  movel([0.295404, -1.335907, -2.579843, -0.796639, 1.570796, 1.866200],accel_mss,speed_ms,0,blend_radius_m)
  movel([0.295412, -1.335943, -2.579820, -0.796627, 1.570796, 1.866208],accel_mss,speed_ms,0,blend_radius_m)
  movel([0.295403, -1.335985, -2.579792, -0.796612, 1.570796, 1.866199],accel_mss,speed_ms,0,blend_radius_m)
  movel([0.295381, -1.336040, -2.579756, -0.796593, 1.570796, 1.866177],accel_mss,speed_ms,0,blend_radius_m)
  movel([0.295349, -1.336095, -2.579721, -0.796574, 1.570796, 1.866145],accel_mss,speed_ms,0,blend_radius_m)
  movel([0.295315, -1.336133, -2.579695, -0.796560, 1.570796, 1.866112],accel_mss,speed_ms,0,blend_radius_m)
  movel([0.295270, -1.336164, -2.579675, -0.796550, 1.570796, 1.866066],accel_mss,speed_ms,0,blend_radius_m)
  movel([0.295209, -1.336190, -2.579659, -0.796541, 1.570796, 1.866006],accel_mss,speed_ms,0,blend_radius_m)
  movel([0.295150, -1.336204, -2.579649, -0.796536, 1.570796, 1.865946],accel_mss,speed_ms,0,blend_radius_m)
  movel([0.294948, -1.336225, -2.579636, -0.796528, 1.570796, 1.865745],accel_mss,speed_ms,0,blend_radius_m)
  movel([0.294564, -1.336243, -2.579624, -0.796522, 1.570796, 1.865360],accel_mss,speed_ms,0,blend_radius_m)
  movel([0.284647, -1.360640, -2.563328, -0.788421, 1.570796, 1.855443],accel_mss,speed_ms,0,blend_radius_m)
  movel([0.280975, -1.369759, -2.557027, -0.785603, 1.570796, 1.851772],accel_mss,speed_ms,0,blend_radius_m)
  movel([0.277925, -1.377354, -2.551691, -0.783344, 1.570796, 1.848721],accel_mss,speed_ms,0,blend_radius_m)
  movel([0.275199, -1.384152, -2.546846, -0.781391, 1.570796, 1.845995],accel_mss,speed_ms,0,blend_radius_m)
  movel([0.275175, -1.384193, -2.546817, -0.781379, 1.570796, 1.845972],accel_mss,speed_ms,0,blend_radius_m)
  movel([0.275139, -1.384229, -2.546791, -0.781369, 1.570796, 1.845936],accel_mss,speed_ms,0,blend_radius_m)
  speed_ms = 0.003
  movel([0.275139, -1.387342, -2.548289, -0.776758, 1.570796, 1.845936],accel_mss,speed_ms,0,blend_radius_m)
  speed_ms = 0.007
  movel([0.275100, -1.387366, -2.548271, -0.776752, 1.570796, 1.845897],accel_mss,speed_ms,0,blend_radius_m)
  movel([0.275061, -1.387375, -2.548265, -0.776749, 1.570796, 1.845858],accel_mss,speed_ms,0,blend_radius_m)
  movel([0.274454, -1.387416, -2.548235, -0.776738, 1.570796, 1.845251],accel_mss,speed_ms,0,blend_radius_m)
  movel([0.273756, -1.387452, -2.548209, -0.776728, 1.570796, 1.844552],accel_mss,speed_ms,0,blend_radius_m)
  movel([0.272946, -1.387481, -2.548189, -0.776720, 1.570796, 1.843742],accel_mss,speed_ms,0,blend_radius_m)
  movel([0.270848, -1.387542, -2.548145, -0.776703, 1.570796, 1.841644],accel_mss,speed_ms,0,blend_radius_m)
  movel([0.270977, -1.387207, -2.548386, -0.776796, 1.570796, 1.841773],accel_mss,speed_ms,0,blend_radius_m)
  movel([0.271720, -1.385272, -2.549778, -0.777339, 1.570796, 1.842517],accel_mss,speed_ms,0,blend_radius_m)
  movel([0.278710, -1.367304, -2.562451, -0.782634, 1.570796, 1.849506],accel_mss,speed_ms,0,blend_radius_m)
  movel([0.285537, -1.349959, -2.574258, -0.788172, 1.570796, 1.856333],accel_mss,speed_ms,0,blend_radius_m)
  movel([0.287626, -1.344699, -2.577757, -0.789933, 1.570796, 1.858423],accel_mss,speed_ms,0,blend_radius_m)
  movel([0.289808, -1.339211, -2.581367, -0.791811, 1.570796, 1.860604],accel_mss,speed_ms,0,blend_radius_m)
  movel([0.289826, -1.339190, -2.581381, -0.791818, 1.570796, 1.860622],accel_mss,speed_ms,0,blend_radius_m)
  movel([0.289853, -1.339171, -2.581393, -0.791825, 1.570796, 1.860650],accel_mss,speed_ms,0,blend_radius_m)
  movel([0.289881, -1.339158, -2.581402, -0.791829, 1.570796, 1.860678],accel_mss,speed_ms,0,blend_radius_m)
  movel([0.289919, -1.339144, -2.581411, -0.791834, 1.570796, 1.860715],accel_mss,speed_ms,0,blend_radius_m)
  movel([0.289955, -1.339137, -2.581415, -0.791836, 1.570796, 1.860751],accel_mss,speed_ms,0,blend_radius_m)
  movel([0.290037, -1.339134, -2.581418, -0.791838, 1.570796, 1.860833],accel_mss,speed_ms,0,blend_radius_m)
  movel([0.294408, -1.339026, -2.581488, -0.791875, 1.570796, 1.865205],accel_mss,speed_ms,0,blend_radius_m)
  movel([0.294728, -1.339025, -2.581489, -0.791875, 1.570796, 1.865524],accel_mss,speed_ms,0,blend_radius_m)
  movel([0.295043, -1.339038, -2.581480, -0.791871, 1.570796, 1.865839],accel_mss,speed_ms,0,blend_radius_m)
  movel([0.295202, -1.339055, -2.581469, -0.791865, 1.570796, 1.865998],accel_mss,speed_ms,0,blend_radius_m)
  movel([0.295351, -1.339089, -2.581447, -0.791853, 1.570796, 1.866147],accel_mss,speed_ms,0,blend_radius_m)
  movel([0.295384, -1.339105, -2.581436, -0.791847, 1.570796, 1.866180],accel_mss,speed_ms,0,blend_radius_m)
  movel([0.295404, -1.339133, -2.581418, -0.791838, 1.570796, 1.866200],accel_mss,speed_ms,0,blend_radius_m)
  movel([0.295412, -1.339168, -2.581395, -0.791826, 1.570796, 1.866208],accel_mss,speed_ms,0,blend_radius_m)
  movel([0.295403, -1.339210, -2.581368, -0.791811, 1.570796, 1.866199],accel_mss,speed_ms,0,blend_radius_m)
  movel([0.295381, -1.339266, -2.581331, -0.791792, 1.570796, 1.866177],accel_mss,speed_ms,0,blend_radius_m)
  movel([0.295349, -1.339320, -2.581296, -0.791773, 1.570796, 1.866145],accel_mss,speed_ms,0,blend_radius_m)
  movel([0.295315, -1.339358, -2.581271, -0.791760, 1.570796, 1.866112],accel_mss,speed_ms,0,blend_radius_m)
  movel([0.295270, -1.339389, -2.581251, -0.791749, 1.570796, 1.866066],accel_mss,speed_ms,0,blend_radius_m)
  movel([0.295209, -1.339415, -2.581234, -0.791740, 1.570796, 1.866006],accel_mss,speed_ms,0,blend_radius_m)
  movel([0.295150, -1.339429, -2.581224, -0.791735, 1.570796, 1.865946],accel_mss,speed_ms,0,blend_radius_m)
  movel([0.294948, -1.339450, -2.581211, -0.791728, 1.570796, 1.865745],accel_mss,speed_ms,0,blend_radius_m)
  movel([0.294564, -1.339468, -2.581199, -0.791722, 1.570796, 1.865360],accel_mss,speed_ms,0,blend_radius_m)
  movel([0.284647, -1.363810, -2.564863, -0.783716, 1.570796, 1.855443],accel_mss,speed_ms,0,blend_radius_m)
  movel([0.280975, -1.372907, -2.558548, -0.780934, 1.570796, 1.851772],accel_mss,speed_ms,0,blend_radius_m)
  movel([0.277925, -1.380483, -2.553200, -0.778706, 1.570796, 1.848721],accel_mss,speed_ms,0,blend_radius_m)
  movel([0.275199, -1.387265, -2.548344, -0.776780, 1.570796, 1.845995],accel_mss,speed_ms,0,blend_radius_m)
  movel([0.275175, -1.387306, -2.548315, -0.776768, 1.570796, 1.845972],accel_mss,speed_ms,0,blend_radius_m)
  movel([0.275139, -1.387342, -2.548289, -0.776758, 1.570796, 1.845936],accel_mss,speed_ms,0,blend_radius_m)
  speed_ms = 0.003
  movel([0.275139, -1.375017, -2.542249, -0.795123, 1.570796, 1.845936],accel_mss,speed_ms,0,blend_radius_m)
  speed_ms = 0.01
  movel([0.275139, -1.351369, -2.529790, -0.831230, 1.570796, 1.845936],accel_mss,speed_ms,0,blend_radius_m)
  movel([0.271209, -1.346627, -2.533019, -0.832743, 1.570796, 1.842006],accel_mss,speed_ms,0,blend_radius_m)
  movel([0.271209, -1.370351, -2.545537, -0.796501, 1.570796, 1.842006],accel_mss,speed_ms,0,blend_radius_m)
  speed_ms = 0.003
  movel([0.271209, -1.379596, -2.550101, -0.782692, 1.570796, 1.842006],accel_mss,speed_ms,0,blend_radius_m)
  speed_ms = 0.007
  movel([0.271117, -1.379629, -2.550077, -0.782683, 1.570796, 1.841914],accel_mss,speed_ms,0,blend_radius_m)
  movel([0.271027, -1.379649, -2.550063, -0.782677, 1.570796, 1.841823],accel_mss,speed_ms,0,blend_radius_m)
  movel([0.270594, -1.379710, -2.550019, -0.782659, 1.570796, 1.841390],accel_mss,speed_ms,0,blend_radius_m)
  movel([0.269882, -1.379801, -2.549955, -0.782633, 1.570796, 1.840679],accel_mss,speed_ms,0,blend_radius_m)
  movel([0.274743, -1.363411, -2.561425, -0.787552, 1.570796, 1.845540],accel_mss,speed_ms,0,blend_radius_m)
  movel([0.279790, -1.346600, -2.572805, -0.792984, 1.570796, 1.850586],accel_mss,speed_ms,0,blend_radius_m)
  movel([0.282065, -1.346298, -2.573006, -0.793085, 1.570796, 1.852861],accel_mss,speed_ms,0,blend_radius_m)
  movel([0.283357, -1.346133, -2.573115, -0.793141, 1.570796, 1.854153],accel_mss,speed_ms,0,blend_radius_m)
  movel([0.283649, -1.346104, -2.573135, -0.793150, 1.570796, 1.854445],accel_mss,speed_ms,0,blend_radius_m)
  movel([0.283936, -1.346085, -2.573147, -0.793157, 1.570796, 1.854732],accel_mss,speed_ms,0,blend_radius_m)
  movel([0.284087, -1.346083, -2.573149, -0.793157, 1.570796, 1.854884],accel_mss,speed_ms,0,blend_radius_m)
  movel([0.284233, -1.346093, -2.573142, -0.793154, 1.570796, 1.855029],accel_mss,speed_ms,0,blend_radius_m)
  movel([0.284260, -1.346103, -2.573135, -0.793151, 1.570796, 1.855057],accel_mss,speed_ms,0,blend_radius_m)
  movel([0.284280, -1.346123, -2.573122, -0.793144, 1.570796, 1.855077],accel_mss,speed_ms,0,blend_radius_m)
  movel([0.284288, -1.346151, -2.573103, -0.793134, 1.570796, 1.855085],accel_mss,speed_ms,0,blend_radius_m)
  movel([0.284283, -1.346184, -2.573082, -0.793124, 1.570796, 1.855079],accel_mss,speed_ms,0,blend_radius_m)
  movel([0.284233, -1.346332, -2.572983, -0.793074, 1.570796, 1.855029],accel_mss,speed_ms,0,blend_radius_m)
  movel([0.282454, -1.350866, -2.569954, -0.791569, 1.570796, 1.853250],accel_mss,speed_ms,0,blend_radius_m)
  movel([0.280494, -1.355873, -2.566576, -0.789940, 1.570796, 1.851291],accel_mss,speed_ms,0,blend_radius_m)
  movel([0.278207, -1.361736, -2.562577, -0.788076, 1.570796, 1.849003],accel_mss,speed_ms,0,blend_radius_m)
  movel([0.275917, -1.367616, -2.558519, -0.786255, 1.570796, 1.846713],accel_mss,speed_ms,0,blend_radius_m)
  movel([0.273935, -1.372723, -2.554954, -0.784711, 1.570796, 1.844731],accel_mss,speed_ms,0,blend_radius_m)
  movel([0.272258, -1.377061, -2.551899, -0.783429, 1.570796, 1.843055],accel_mss,speed_ms,0,blend_radius_m)
  movel([0.271919, -1.377934, -2.551281, -0.783175, 1.570796, 1.842716],accel_mss,speed_ms,0,blend_radius_m)
  movel([0.271351, -1.379441, -2.550211, -0.782737, 1.570796, 1.842148],accel_mss,speed_ms,0,blend_radius_m)
  movel([0.271312, -1.379512, -2.550160, -0.782717, 1.570796, 1.842108],accel_mss,speed_ms,0,blend_radius_m)
  movel([0.271281, -1.379546, -2.550136, -0.782707, 1.570796, 1.842078],accel_mss,speed_ms,0,blend_radius_m)
  movel([0.271248, -1.379574, -2.550116, -0.782699, 1.570796, 1.842044],accel_mss,speed_ms,0,blend_radius_m)
  movel([0.271209, -1.379596, -2.550101, -0.782692, 1.570796, 1.842006],accel_mss,speed_ms,0,blend_radius_m)
  speed_ms = 0.003
  movel([0.271209, -1.382720, -2.551606, -0.778063, 1.570796, 1.842006],accel_mss,speed_ms,0,blend_radius_m)
  speed_ms = 0.007
  movel([0.271117, -1.382753, -2.551582, -0.778054, 1.570796, 1.841914],accel_mss,speed_ms,0,blend_radius_m)
  movel([0.271027, -1.382773, -2.551568, -0.778048, 1.570796, 1.841823],accel_mss,speed_ms,0,blend_radius_m)
  movel([0.270594, -1.382834, -2.551524, -0.778031, 1.570796, 1.841390],accel_mss,speed_ms,0,blend_radius_m)
  movel([0.269882, -1.382924, -2.551460, -0.778005, 1.570796, 1.840679],accel_mss,speed_ms,0,blend_radius_m)
  movel([0.274743, -1.366574, -2.562956, -0.782858, 1.570796, 1.845540],accel_mss,speed_ms,0,blend_radius_m)
  movel([0.279790, -1.349802, -2.574363, -0.788224, 1.570796, 1.850586],accel_mss,speed_ms,0,blend_radius_m)
  movel([0.282065, -1.349501, -2.574564, -0.788324, 1.570796, 1.852861],accel_mss,speed_ms,0,blend_radius_m)
  movel([0.283357, -1.349336, -2.574674, -0.788379, 1.570796, 1.854153],accel_mss,speed_ms,0,blend_radius_m)
  movel([0.283649, -1.349307, -2.574694, -0.788388, 1.570796, 1.854445],accel_mss,speed_ms,0,blend_radius_m)
  movel([0.283936, -1.349288, -2.574707, -0.788395, 1.570796, 1.854732],accel_mss,speed_ms,0,blend_radius_m)
  movel([0.284087, -1.349286, -2.574708, -0.788395, 1.570796, 1.854884],accel_mss,speed_ms,0,blend_radius_m)
  movel([0.284233, -1.349296, -2.574701, -0.788392, 1.570796, 1.855029],accel_mss,speed_ms,0,blend_radius_m)
  movel([0.284260, -1.349306, -2.574694, -0.788389, 1.570796, 1.855057],accel_mss,speed_ms,0,blend_radius_m)
  movel([0.284280, -1.349326, -2.574681, -0.788382, 1.570796, 1.855077],accel_mss,speed_ms,0,blend_radius_m)
  movel([0.284288, -1.349354, -2.574662, -0.788373, 1.570796, 1.855085],accel_mss,speed_ms,0,blend_radius_m)
  movel([0.284283, -1.349386, -2.574641, -0.788362, 1.570796, 1.855079],accel_mss,speed_ms,0,blend_radius_m)
  movel([0.284233, -1.349534, -2.574542, -0.788313, 1.570796, 1.855029],accel_mss,speed_ms,0,blend_radius_m)
  movel([0.282454, -1.354058, -2.571505, -0.786826, 1.570796, 1.853250],accel_mss,speed_ms,0,blend_radius_m)
  movel([0.280494, -1.359054, -2.568119, -0.785216, 1.570796, 1.851291],accel_mss,speed_ms,0,blend_radius_m)
  movel([0.278207, -1.364903, -2.564110, -0.783376, 1.570796, 1.849003],accel_mss,speed_ms,0,blend_radius_m)
  movel([0.275917, -1.370769, -2.560043, -0.781578, 1.570796, 1.846713],accel_mss,speed_ms,0,blend_radius_m)
  movel([0.273935, -1.375864, -2.556470, -0.780055, 1.570796, 1.844731],accel_mss,speed_ms,0,blend_radius_m)
  movel([0.272258, -1.380191, -2.553408, -0.778790, 1.570796, 1.843055],accel_mss,speed_ms,0,blend_radius_m)
  movel([0.271919, -1.381062, -2.552788, -0.778539, 1.570796, 1.842716],accel_mss,speed_ms,0,blend_radius_m)
  movel([0.271351, -1.382565, -2.551716, -0.778107, 1.570796, 1.842148],accel_mss,speed_ms,0,blend_radius_m)
  movel([0.271312, -1.382637, -2.551665, -0.778087, 1.570796, 1.842108],accel_mss,speed_ms,0,blend_radius_m)
  movel([0.271281, -1.382670, -2.551641, -0.778077, 1.570796, 1.842078],accel_mss,speed_ms,0,blend_radius_m)
  movel([0.271248, -1.382698, -2.551621, -0.778069, 1.570796, 1.842044],accel_mss,speed_ms,0,blend_radius_m)
  movel([0.271209, -1.382720, -2.551606, -0.778063, 1.570796, 1.842006],accel_mss,speed_ms,0,blend_radius_m)
  speed_ms = 0.003
  movel([0.271209, -1.370351, -2.545537, -0.796501, 1.570796, 1.842006],accel_mss,speed_ms,0,blend_radius_m)
  speed_ms = 0.01
  movel([0.271209, -1.346627, -2.533019, -0.832743, 1.570796, 1.842006],accel_mss,speed_ms,0,blend_radius_m)
  movel([0.283720, -1.297614, -2.564685, -0.850089, 1.570796, 1.854516],accel_mss,speed_ms,0,blend_radius_m)
  movel([0.283720, -1.322065, -2.577821, -0.812503, 1.570796, 1.854516],accel_mss,speed_ms,0,blend_radius_m)
  speed_ms = 0.003
  movel([0.283720, -1.331626, -2.582617, -0.798146, 1.570796, 1.854516],accel_mss,speed_ms,0,blend_radius_m)
  speed_ms = 0.007
  movel([0.283274, -1.331697, -2.582572, -0.798121, 1.570796, 1.854071],accel_mss,speed_ms,0,blend_radius_m)
  movel([0.282766, -1.331776, -2.582521, -0.798093, 1.570796, 1.853563],accel_mss,speed_ms,0,blend_radius_m)
  movel([0.282165, -1.331861, -2.582466, -0.798062, 1.570796, 1.852961],accel_mss,speed_ms,0,blend_radius_m)
  movel([0.280602, -1.332079, -2.582325, -0.797985, 1.570796, 1.851398],accel_mss,speed_ms,0,blend_radius_m)
  movel([0.280741, -1.331617, -2.582623, -0.798149, 1.570796, 1.851537],accel_mss,speed_ms,0,blend_radius_m)
  movel([0.280880, -1.331154, -2.582922, -0.798313, 1.570796, 1.851676],accel_mss,speed_ms,0,blend_radius_m)
  movel([0.282316, -1.331363, -2.582787, -0.798239, 1.570796, 1.853112],accel_mss,speed_ms,0,blend_radius_m)
  movel([0.282867, -1.331445, -2.582734, -0.798210, 1.570796, 1.853663],accel_mss,speed_ms,0,blend_radius_m)
  movel([0.283328, -1.331519, -2.582686, -0.798184, 1.570796, 1.854125],accel_mss,speed_ms,0,blend_radius_m)
  movel([0.283733, -1.331590, -2.582641, -0.798158, 1.570796, 1.854530],accel_mss,speed_ms,0,blend_radius_m)
  movel([0.283741, -1.331598, -2.582635, -0.798156, 1.570796, 1.854537],accel_mss,speed_ms,0,blend_radius_m)
  movel([0.283739, -1.331610, -2.582628, -0.798151, 1.570796, 1.854536],accel_mss,speed_ms,0,blend_radius_m)
  movel([0.283720, -1.331626, -2.582617, -0.798146, 1.570796, 1.854516],accel_mss,speed_ms,0,blend_radius_m)
  speed_ms = 0.003
  movel([0.283720, -1.334861, -2.584200, -0.793328, 1.570796, 1.854516],accel_mss,speed_ms,0,blend_radius_m)
  speed_ms = 0.007
  movel([0.283274, -1.334931, -2.584154, -0.793303, 1.570796, 1.854071],accel_mss,speed_ms,0,blend_radius_m)
  movel([0.282766, -1.335010, -2.584103, -0.793275, 1.570796, 1.853563],accel_mss,speed_ms,0,blend_radius_m)
  movel([0.282165, -1.335096, -2.584048, -0.793245, 1.570796, 1.852961],accel_mss,speed_ms,0,blend_radius_m)
  movel([0.280602, -1.335313, -2.583907, -0.793169, 1.570796, 1.851398],accel_mss,speed_ms,0,blend_radius_m)
  movel([0.280741, -1.334852, -2.584206, -0.793331, 1.570796, 1.851537],accel_mss,speed_ms,0,blend_radius_m)
  movel([0.280880, -1.334390, -2.584505, -0.793494, 1.570796, 1.851676],accel_mss,speed_ms,0,blend_radius_m)
  movel([0.282316, -1.334598, -2.584370, -0.793420, 1.570796, 1.853112],accel_mss,speed_ms,0,blend_radius_m)
  movel([0.282867, -1.334681, -2.584317, -0.793391, 1.570796, 1.853663],accel_mss,speed_ms,0,blend_radius_m)
  movel([0.283328, -1.334754, -2.584269, -0.793365, 1.570796, 1.854125],accel_mss,speed_ms,0,blend_radius_m)
  movel([0.283733, -1.334825, -2.584223, -0.793341, 1.570796, 1.854530],accel_mss,speed_ms,0,blend_radius_m)
  movel([0.283741, -1.334833, -2.584218, -0.793338, 1.570796, 1.854537],accel_mss,speed_ms,0,blend_radius_m)
  movel([0.283739, -1.334845, -2.584211, -0.793334, 1.570796, 1.854536],accel_mss,speed_ms,0,blend_radius_m)
  movel([0.283720, -1.334861, -2.584200, -0.793328, 1.570796, 1.854516],accel_mss,speed_ms,0,blend_radius_m)
  speed_ms = 0.003
  movel([0.283720, -1.322065, -2.577821, -0.812503, 1.570796, 1.854516],accel_mss,speed_ms,0,blend_radius_m)
  speed_ms = 0.01
  movel([0.283720, -1.297614, -2.564685, -0.850089, 1.570796, 1.854516],accel_mss,speed_ms,0,blend_radius_m)
  movel([0.283763, -1.295871, -2.565756, -0.850763, 1.570796, 1.854559],accel_mss,speed_ms,0,blend_radius_m)
  movel([0.283763, -1.320346, -2.578913, -0.813130, 1.570796, 1.854559],accel_mss,speed_ms,0,blend_radius_m)
  speed_ms = 0.003
  movel([0.283763, -1.329917, -2.583718, -0.798754, 1.570796, 1.854559],accel_mss,speed_ms,0,blend_radius_m)
  speed_ms = 0.007
  movel([0.283665, -1.329924, -2.583714, -0.798751, 1.570796, 1.854461],accel_mss,speed_ms,0,blend_radius_m)
  movel([0.283573, -1.329918, -2.583718, -0.798754, 1.570796, 1.854369],accel_mss,speed_ms,0,blend_radius_m)
  movel([0.267806, -1.327695, -2.585144, -0.799550, 1.570796, 1.838602],accel_mss,speed_ms,0,blend_radius_m)
  movel([0.251809, -1.325748, -2.586388, -0.800254, 1.570796, 1.822605],accel_mss,speed_ms,0,blend_radius_m)
  movel([0.251761, -1.325735, -2.586396, -0.800258, 1.570796, 1.822557],accel_mss,speed_ms,0,blend_radius_m)
  movel([0.251724, -1.325709, -2.586412, -0.800268, 1.570796, 1.822521],accel_mss,speed_ms,0,blend_radius_m)
  movel([0.251715, -1.325681, -2.586430, -0.800278, 1.570796, 1.822511],accel_mss,speed_ms,0,blend_radius_m)
  movel([0.251725, -1.325645, -2.586453, -0.800291, 1.570796, 1.822521],accel_mss,speed_ms,0,blend_radius_m)
  movel([0.254190, -1.320979, -2.589413, -0.801998, 1.570796, 1.824987],accel_mss,speed_ms,0,blend_radius_m)
  movel([0.256668, -1.316306, -2.592348, -0.803735, 1.570796, 1.827464],accel_mss,speed_ms,0,blend_radius_m)
  movel([0.256713, -1.316240, -2.592389, -0.803760, 1.570796, 1.827509],accel_mss,speed_ms,0,blend_radius_m)
  movel([0.256772, -1.316177, -2.592429, -0.803784, 1.570796, 1.827569],accel_mss,speed_ms,0,blend_radius_m)
  movel([0.256793, -1.316164, -2.592437, -0.803789, 1.570796, 1.827589],accel_mss,speed_ms,0,blend_radius_m)
  movel([0.256813, -1.316160, -2.592439, -0.803790, 1.570796, 1.827610],accel_mss,speed_ms,0,blend_radius_m)
  movel([0.257759, -1.316208, -2.592409, -0.803772, 1.570796, 1.828555],accel_mss,speed_ms,0,blend_radius_m)
  movel([0.258816, -1.316268, -2.592371, -0.803750, 1.570796, 1.829612],accel_mss,speed_ms,0,blend_radius_m)
  movel([0.260062, -1.316349, -2.592321, -0.803719, 1.570796, 1.830859],accel_mss,speed_ms,0,blend_radius_m)
  movel([0.263935, -1.316628, -2.592146, -0.803615, 1.570796, 1.834731],accel_mss,speed_ms,0,blend_radius_m)
  movel([0.267792, -1.316934, -2.591955, -0.803500, 1.570796, 1.838588],accel_mss,speed_ms,0,blend_radius_m)
  movel([0.269155, -1.317054, -2.591880, -0.803455, 1.570796, 1.839952],accel_mss,speed_ms,0,blend_radius_m)
  movel([0.270512, -1.317186, -2.591797, -0.803406, 1.570796, 1.841308],accel_mss,speed_ms,0,blend_radius_m)
  movel([0.271861, -1.317333, -2.591705, -0.803351, 1.570796, 1.842657],accel_mss,speed_ms,0,blend_radius_m)
  movel([0.272781, -1.317446, -2.591634, -0.803309, 1.570796, 1.843577],accel_mss,speed_ms,0,blend_radius_m)
  movel([0.273693, -1.317576, -2.591553, -0.803260, 1.570796, 1.844489],accel_mss,speed_ms,0,blend_radius_m)
  movel([0.274595, -1.317721, -2.591462, -0.803206, 1.570796, 1.845392],accel_mss,speed_ms,0,blend_radius_m)
  movel([0.275414, -1.317867, -2.591370, -0.803152, 1.570796, 1.846211],accel_mss,speed_ms,0,blend_radius_m)
  movel([0.276222, -1.318035, -2.591265, -0.803089, 1.570796, 1.847018],accel_mss,speed_ms,0,blend_radius_m)
  movel([0.277016, -1.318219, -2.591150, -0.803021, 1.570796, 1.847813],accel_mss,speed_ms,0,blend_radius_m)
  movel([0.277714, -1.318399, -2.591036, -0.802953, 1.570796, 1.848511],accel_mss,speed_ms,0,blend_radius_m)
  movel([0.278399, -1.318598, -2.590911, -0.802879, 1.570796, 1.849196],accel_mss,speed_ms,0,blend_radius_m)
  movel([0.279071, -1.318816, -2.590774, -0.802798, 1.570796, 1.849867],accel_mss,speed_ms,0,blend_radius_m)
  movel([0.279730, -1.319051, -2.590627, -0.802711, 1.570796, 1.850526],accel_mss,speed_ms,0,blend_radius_m)
  movel([0.280376, -1.319301, -2.590469, -0.802618, 1.570796, 1.851173],accel_mss,speed_ms,0,blend_radius_m)
  movel([0.281010, -1.319571, -2.590300, -0.802518, 1.570796, 1.851806],accel_mss,speed_ms,0,blend_radius_m)
  movel([0.281379, -1.319745, -2.590190, -0.802454, 1.570796, 1.852176],accel_mss,speed_ms,0,blend_radius_m)
  movel([0.281738, -1.319934, -2.590071, -0.802384, 1.570796, 1.852534],accel_mss,speed_ms,0,blend_radius_m)
  movel([0.282081, -1.320138, -2.589943, -0.802308, 1.570796, 1.852878],accel_mss,speed_ms,0,blend_radius_m)
  movel([0.282417, -1.320353, -2.589807, -0.802229, 1.570796, 1.853213],accel_mss,speed_ms,0,blend_radius_m)
  movel([0.282735, -1.320585, -2.589661, -0.802143, 1.570796, 1.853531],accel_mss,speed_ms,0,blend_radius_m)
  movel([0.283041, -1.320830, -2.589506, -0.802052, 1.570796, 1.853838],accel_mss,speed_ms,0,blend_radius_m)
  movel([0.283334, -1.321089, -2.589343, -0.801957, 1.570796, 1.854130],accel_mss,speed_ms,0,blend_radius_m)
  movel([0.283610, -1.321359, -2.589172, -0.801857, 1.570796, 1.854407],accel_mss,speed_ms,0,blend_radius_m)
  movel([0.283835, -1.321600, -2.589020, -0.801769, 1.570796, 1.854632],accel_mss,speed_ms,0,blend_radius_m)
  movel([0.284041, -1.321857, -2.588858, -0.801674, 1.570796, 1.854837],accel_mss,speed_ms,0,blend_radius_m)
  movel([0.284233, -1.322123, -2.588690, -0.801577, 1.570796, 1.855030],accel_mss,speed_ms,0,blend_radius_m)
  movel([0.284407, -1.322403, -2.588512, -0.801474, 1.570796, 1.855203],accel_mss,speed_ms,0,blend_radius_m)
  movel([0.284568, -1.322694, -2.588328, -0.801367, 1.570796, 1.855364],accel_mss,speed_ms,0,blend_radius_m)
  movel([0.284710, -1.322997, -2.588136, -0.801256, 1.570796, 1.855506],accel_mss,speed_ms,0,blend_radius_m)
  movel([0.284835, -1.323310, -2.587938, -0.801141, 1.570796, 1.855631],accel_mss,speed_ms,0,blend_radius_m)
  movel([0.284944, -1.323634, -2.587732, -0.801023, 1.570796, 1.855740],accel_mss,speed_ms,0,blend_radius_m)
  movel([0.285032, -1.323956, -2.587528, -0.800906, 1.570796, 1.855828],accel_mss,speed_ms,0,blend_radius_m)
  movel([0.285100, -1.324285, -2.587319, -0.800785, 1.570796, 1.855897],accel_mss,speed_ms,0,blend_radius_m)
  movel([0.285151, -1.324626, -2.587102, -0.800661, 1.570796, 1.855947],accel_mss,speed_ms,0,blend_radius_m)
  movel([0.285182, -1.324974, -2.586880, -0.800535, 1.570796, 1.855979],accel_mss,speed_ms,0,blend_radius_m)
  movel([0.285194, -1.325332, -2.586653, -0.800405, 1.570796, 1.855990],accel_mss,speed_ms,0,blend_radius_m)
  movel([0.285186, -1.325696, -2.586420, -0.800272, 1.570796, 1.855982],accel_mss,speed_ms,0,blend_radius_m)
  movel([0.285163, -1.326065, -2.586185, -0.800139, 1.570796, 1.855959],accel_mss,speed_ms,0,blend_radius_m)
  movel([0.285118, -1.326442, -2.585945, -0.800002, 1.570796, 1.855914],accel_mss,speed_ms,0,blend_radius_m)
  movel([0.285089, -1.326615, -2.585834, -0.799940, 1.570796, 1.855885],accel_mss,speed_ms,0,blend_radius_m)
  movel([0.285048, -1.326789, -2.585723, -0.799877, 1.570796, 1.855844],accel_mss,speed_ms,0,blend_radius_m)
  movel([0.284996, -1.326967, -2.585609, -0.799813, 1.570796, 1.855792],accel_mss,speed_ms,0,blend_radius_m)
  movel([0.284808, -1.327550, -2.585236, -0.799602, 1.570796, 1.855605],accel_mss,speed_ms,0,blend_radius_m)
  movel([0.284614, -1.328133, -2.584863, -0.799393, 1.570796, 1.855410],accel_mss,speed_ms,0,blend_radius_m)
  movel([0.284200, -1.329332, -2.584094, -0.798963, 1.570796, 1.854997],accel_mss,speed_ms,0,blend_radius_m)
  movel([0.284152, -1.329451, -2.584018, -0.798920, 1.570796, 1.854948],accel_mss,speed_ms,0,blend_radius_m)
  movel([0.284092, -1.329568, -2.583943, -0.798879, 1.570796, 1.854889],accel_mss,speed_ms,0,blend_radius_m)
  movel([0.284020, -1.329686, -2.583867, -0.798836, 1.570796, 1.854817],accel_mss,speed_ms,0,blend_radius_m)
  movel([0.283957, -1.329768, -2.583814, -0.798807, 1.570796, 1.854753],accel_mss,speed_ms,0,blend_radius_m)
  movel([0.283884, -1.329843, -2.583766, -0.798780, 1.570796, 1.854680],accel_mss,speed_ms,0,blend_radius_m)
  movel([0.283815, -1.329896, -2.583732, -0.798761, 1.570796, 1.854611],accel_mss,speed_ms,0,blend_radius_m)
  movel([0.283789, -1.329909, -2.583723, -0.798757, 1.570796, 1.854586],accel_mss,speed_ms,0,blend_radius_m)
  movel([0.283763, -1.329917, -2.583718, -0.798754, 1.570796, 1.854559],accel_mss,speed_ms,0,blend_radius_m)
  speed_ms = 0.003
  movel([0.283763, -1.333156, -2.585304, -0.793930, 1.570796, 1.854559],accel_mss,speed_ms,0,blend_radius_m)
  speed_ms = 0.007
  movel([0.283665, -1.333162, -2.585299, -0.793927, 1.570796, 1.854461],accel_mss,speed_ms,0,blend_radius_m)
  movel([0.283573, -1.333157, -2.585303, -0.793929, 1.570796, 1.854369],accel_mss,speed_ms,0,blend_radius_m)
  movel([0.267806, -1.330938, -2.586733, -0.794718, 1.570796, 1.838602],accel_mss,speed_ms,0,blend_radius_m)
  movel([0.251809, -1.328995, -2.587980, -0.795414, 1.570796, 1.822605],accel_mss,speed_ms,0,blend_radius_m)
  movel([0.251761, -1.328983, -2.587988, -0.795418, 1.570796, 1.822557],accel_mss,speed_ms,0,blend_radius_m)
  movel([0.251724, -1.328957, -2.588005, -0.795428, 1.570796, 1.822521],accel_mss,speed_ms,0,blend_radius_m)
  movel([0.251715, -1.328929, -2.588023, -0.795438, 1.570796, 1.822511],accel_mss,speed_ms,0,blend_radius_m)
  movel([0.251725, -1.328893, -2.588046, -0.795451, 1.570796, 1.822521],accel_mss,speed_ms,0,blend_radius_m)
  movel([0.254190, -1.324237, -2.591013, -0.797140, 1.570796, 1.824987],accel_mss,speed_ms,0,blend_radius_m)
  movel([0.256668, -1.319574, -2.593956, -0.798860, 1.570796, 1.827464],accel_mss,speed_ms,0,blend_radius_m)
  movel([0.256713, -1.319508, -2.593997, -0.798884, 1.570796, 1.827509],accel_mss,speed_ms,0,blend_radius_m)
  movel([0.256772, -1.319445, -2.594037, -0.798908, 1.570796, 1.827569],accel_mss,speed_ms,0,blend_radius_m)
  movel([0.256793, -1.319432, -2.594045, -0.798913, 1.570796, 1.827589],accel_mss,speed_ms,0,blend_radius_m)
  movel([0.256813, -1.319428, -2.594047, -0.798914, 1.570796, 1.827610],accel_mss,speed_ms,0,blend_radius_m)
  movel([0.257759, -1.319476, -2.594017, -0.798896, 1.570796, 1.828555],accel_mss,speed_ms,0,blend_radius_m)
  movel([0.258816, -1.319536, -2.593979, -0.798874, 1.570796, 1.829612],accel_mss,speed_ms,0,blend_radius_m)
  movel([0.260062, -1.319616, -2.593929, -0.798844, 1.570796, 1.830859],accel_mss,speed_ms,0,blend_radius_m)
  movel([0.263935, -1.319895, -2.593754, -0.798740, 1.570796, 1.834731],accel_mss,speed_ms,0,blend_radius_m)
  movel([0.267792, -1.320200, -2.593562, -0.798627, 1.570796, 1.838588],accel_mss,speed_ms,0,blend_radius_m)
  movel([0.269155, -1.320320, -2.593486, -0.798582, 1.570796, 1.839952],accel_mss,speed_ms,0,blend_radius_m)
  movel([0.270512, -1.320452, -2.593403, -0.798533, 1.570796, 1.841308],accel_mss,speed_ms,0,blend_radius_m)
  movel([0.271861, -1.320599, -2.593311, -0.798479, 1.570796, 1.842657],accel_mss,speed_ms,0,blend_radius_m)
  movel([0.272781, -1.320711, -2.593240, -0.798438, 1.570796, 1.843577],accel_mss,speed_ms,0,blend_radius_m)
  movel([0.273693, -1.320841, -2.593158, -0.798389, 1.570796, 1.844489],accel_mss,speed_ms,0,blend_radius_m)
  movel([0.274595, -1.320986, -2.593068, -0.798336, 1.570796, 1.845392],accel_mss,speed_ms,0,blend_radius_m)
  movel([0.275414, -1.321132, -2.592975, -0.798282, 1.570796, 1.846211],accel_mss,speed_ms,0,blend_radius_m)
  movel([0.276222, -1.321299, -2.592870, -0.798220, 1.570796, 1.847018],accel_mss,speed_ms,0,blend_radius_m)
  movel([0.277016, -1.321483, -2.592754, -0.798152, 1.570796, 1.847813],accel_mss,speed_ms,0,blend_radius_m)
  movel([0.277714, -1.321663, -2.592641, -0.798086, 1.570796, 1.848511],accel_mss,speed_ms,0,blend_radius_m)
  movel([0.278399, -1.321861, -2.592515, -0.798012, 1.570796, 1.849196],accel_mss,speed_ms,0,blend_radius_m)
  movel([0.279071, -1.322079, -2.592378, -0.797932, 1.570796, 1.849867],accel_mss,speed_ms,0,blend_radius_m)
  movel([0.279730, -1.322313, -2.592230, -0.797846, 1.570796, 1.850526],accel_mss,speed_ms,0,blend_radius_m)
  movel([0.280376, -1.322563, -2.592072, -0.797754, 1.570796, 1.851173],accel_mss,speed_ms,0,blend_radius_m)
  movel([0.281010, -1.322831, -2.591903, -0.797655, 1.570796, 1.851806],accel_mss,speed_ms,0,blend_radius_m)
  movel([0.281379, -1.323006, -2.591792, -0.797591, 1.570796, 1.852176],accel_mss,speed_ms,0,blend_radius_m)
  movel([0.281738, -1.323194, -2.591673, -0.797522, 1.570796, 1.852534],accel_mss,speed_ms,0,blend_radius_m)
  movel([0.282081, -1.323398, -2.591544, -0.797447, 1.570796, 1.852878],accel_mss,speed_ms,0,blend_radius_m)
  movel([0.282417, -1.323613, -2.591408, -0.797368, 1.570796, 1.853213],accel_mss,speed_ms,0,blend_radius_m)
  movel([0.282735, -1.323844, -2.591262, -0.797283, 1.570796, 1.853531],accel_mss,speed_ms,0,blend_radius_m)
  movel([0.283041, -1.324088, -2.591107, -0.797194, 1.570796, 1.853838],accel_mss,speed_ms,0,blend_radius_m)
  movel([0.283334, -1.324347, -2.590943, -0.797099, 1.570796, 1.854130],accel_mss,speed_ms,0,blend_radius_m)
  movel([0.283610, -1.324616, -2.590772, -0.797001, 1.570796, 1.854407],accel_mss,speed_ms,0,blend_radius_m)
  movel([0.283835, -1.324856, -2.590620, -0.796913, 1.570796, 1.854632],accel_mss,speed_ms,0,blend_radius_m)
  movel([0.284041, -1.325113, -2.590457, -0.796820, 1.570796, 1.854837],accel_mss,speed_ms,0,blend_radius_m)
  movel([0.284233, -1.325378, -2.590288, -0.796723, 1.570796, 1.855030],accel_mss,speed_ms,0,blend_radius_m)
  movel([0.284407, -1.325658, -2.590110, -0.796621, 1.570796, 1.855203],accel_mss,speed_ms,0,blend_radius_m)
  movel([0.284568, -1.325949, -2.589925, -0.796515, 1.570796, 1.855364],accel_mss,speed_ms,0,blend_radius_m)
  movel([0.284710, -1.326251, -2.589733, -0.796405, 1.570796, 1.855506],accel_mss,speed_ms,0,blend_radius_m)
  movel([0.284835, -1.326563, -2.589534, -0.796292, 1.570796, 1.855631],accel_mss,speed_ms,0,blend_radius_m)
  movel([0.284944, -1.326886, -2.589328, -0.796175, 1.570796, 1.855740],accel_mss,speed_ms,0,blend_radius_m)
  movel([0.285032, -1.327207, -2.589123, -0.796059, 1.570796, 1.855828],accel_mss,speed_ms,0,blend_radius_m)
  movel([0.285100, -1.327536, -2.588913, -0.795940, 1.570796, 1.855897],accel_mss,speed_ms,0,blend_radius_m)
  movel([0.285151, -1.327876, -2.588696, -0.795817, 1.570796, 1.855947],accel_mss,speed_ms,0,blend_radius_m)
  movel([0.285182, -1.328223, -2.588474, -0.795692, 1.570796, 1.855979],accel_mss,speed_ms,0,blend_radius_m)
  movel([0.285194, -1.328580, -2.588246, -0.795563, 1.570796, 1.855990],accel_mss,speed_ms,0,blend_radius_m)
  movel([0.285186, -1.328944, -2.588013, -0.795432, 1.570796, 1.855982],accel_mss,speed_ms,0,blend_radius_m)
  movel([0.285163, -1.329312, -2.587777, -0.795300, 1.570796, 1.855959],accel_mss,speed_ms,0,blend_radius_m)
  movel([0.285118, -1.329688, -2.587536, -0.795165, 1.570796, 1.855914],accel_mss,speed_ms,0,blend_radius_m)
  movel([0.285089, -1.329861, -2.587425, -0.795103, 1.570796, 1.855885],accel_mss,speed_ms,0,blend_radius_m)
  movel([0.285048, -1.330035, -2.587314, -0.795041, 1.570796, 1.855844],accel_mss,speed_ms,0,blend_radius_m)
  movel([0.284996, -1.330213, -2.587199, -0.794977, 1.570796, 1.855792],accel_mss,speed_ms,0,blend_radius_m)
  movel([0.284808, -1.330794, -2.586826, -0.794769, 1.570796, 1.855605],accel_mss,speed_ms,0,blend_radius_m)
  movel([0.284614, -1.331376, -2.586451, -0.794562, 1.570796, 1.855410],accel_mss,speed_ms,0,blend_radius_m)
  movel([0.284200, -1.332572, -2.585681, -0.794137, 1.570796, 1.854997],accel_mss,speed_ms,0,blend_radius_m)
  movel([0.284152, -1.332691, -2.585604, -0.794094, 1.570796, 1.854948],accel_mss,speed_ms,0,blend_radius_m)
  movel([0.284092, -1.332807, -2.585529, -0.794053, 1.570796, 1.854889],accel_mss,speed_ms,0,blend_radius_m)
  movel([0.284020, -1.332925, -2.585453, -0.794011, 1.570796, 1.854817],accel_mss,speed_ms,0,blend_radius_m)
  movel([0.283957, -1.333007, -2.585400, -0.793982, 1.570796, 1.854753],accel_mss,speed_ms,0,blend_radius_m)
  movel([0.283884, -1.333082, -2.585352, -0.793956, 1.570796, 1.854680],accel_mss,speed_ms,0,blend_radius_m)
  movel([0.283815, -1.333135, -2.585317, -0.793937, 1.570796, 1.854611],accel_mss,speed_ms,0,blend_radius_m)
  movel([0.283789, -1.333147, -2.585309, -0.793932, 1.570796, 1.854586],accel_mss,speed_ms,0,blend_radius_m)
  movel([0.283763, -1.333156, -2.585304, -0.793930, 1.570796, 1.854559],accel_mss,speed_ms,0,blend_radius_m)
  speed_ms = 0.003
  movel([0.283763, -1.320346, -2.578913, -0.813130, 1.570796, 1.854559],accel_mss,speed_ms,0,blend_radius_m)
  speed_ms = 0.01
  movel([0.283763, -1.295871, -2.565756, -0.850763, 1.570796, 1.854559],accel_mss,speed_ms,0,blend_radius_m)
  movel([0.282293, -1.299239, -2.563684, -0.849465, 1.570796, 1.853089],accel_mss,speed_ms,0,blend_radius_m)
  movel([0.282293, -1.323668, -2.576799, -0.811922, 1.570796, 1.853089],accel_mss,speed_ms,0,blend_radius_m)
  speed_ms = 0.003
  movel([0.282293, -1.333219, -2.581588, -0.797582, 1.570796, 1.853089],accel_mss,speed_ms,0,blend_radius_m)
  speed_ms = 0.007
  movel([0.281918, -1.334455, -2.580786, -0.797147, 1.570796, 1.852714],accel_mss,speed_ms,0,blend_radius_m)
  movel([0.281544, -1.335690, -2.579984, -0.796715, 1.570796, 1.852341],accel_mss,speed_ms,0,blend_radius_m)
  movel([0.278441, -1.336188, -2.579660, -0.796541, 1.570796, 1.849238],accel_mss,speed_ms,0,blend_radius_m)
  movel([0.276251, -1.336569, -2.579411, -0.796409, 1.570796, 1.847047],accel_mss,speed_ms,0,blend_radius_m)
  movel([0.275394, -1.336738, -2.579301, -0.796350, 1.570796, 1.846190],accel_mss,speed_ms,0,blend_radius_m)
  movel([0.274530, -1.336932, -2.579175, -0.796282, 1.570796, 1.845326],accel_mss,speed_ms,0,blend_radius_m)
  movel([0.273708, -1.337136, -2.579041, -0.796211, 1.570796, 1.844505],accel_mss,speed_ms,0,blend_radius_m)
  movel([0.272883, -1.337362, -2.578894, -0.796133, 1.570796, 1.843679],accel_mss,speed_ms,0,blend_radius_m)
  movel([0.270940, -1.337952, -2.578508, -0.795928, 1.570796, 1.841736],accel_mss,speed_ms,0,blend_radius_m)
  movel([0.269926, -1.338289, -2.578288, -0.795812, 1.570796, 1.840722],accel_mss,speed_ms,0,blend_radius_m)
  movel([0.268912, -1.338651, -2.578052, -0.795687, 1.570796, 1.839708],accel_mss,speed_ms,0,blend_radius_m)
  movel([0.267897, -1.339034, -2.577801, -0.795555, 1.570796, 1.838694],accel_mss,speed_ms,0,blend_radius_m)
  movel([0.266884, -1.339440, -2.577535, -0.795415, 1.570796, 1.837680],accel_mss,speed_ms,0,blend_radius_m)
  movel([0.265880, -1.339865, -2.577256, -0.795268, 1.570796, 1.836676],accel_mss,speed_ms,0,blend_radius_m)
  movel([0.264877, -1.340313, -2.576961, -0.795114, 1.570796, 1.835673],accel_mss,speed_ms,0,blend_radius_m)
  movel([0.263878, -1.340784, -2.576652, -0.794953, 1.570796, 1.834675],accel_mss,speed_ms,0,blend_radius_m)
  movel([0.262881, -1.341275, -2.576329, -0.794785, 1.570796, 1.833678],accel_mss,speed_ms,0,blend_radius_m)
  movel([0.261910, -1.341780, -2.575996, -0.794613, 1.570796, 1.832706],accel_mss,speed_ms,0,blend_radius_m)
  movel([0.260943, -1.342306, -2.575650, -0.794434, 1.570796, 1.831739],accel_mss,speed_ms,0,blend_radius_m)
  movel([0.259983, -1.342850, -2.575290, -0.794248, 1.570796, 1.830780],accel_mss,speed_ms,0,blend_radius_m)
  movel([0.259028, -1.343417, -2.574916, -0.794056, 1.570796, 1.829824],accel_mss,speed_ms,0,blend_radius_m)
  movel([0.258111, -1.343985, -2.574540, -0.793864, 1.570796, 1.828907],accel_mss,speed_ms,0,blend_radius_m)
  movel([0.257201, -1.344573, -2.574150, -0.793665, 1.570796, 1.827997],accel_mss,speed_ms,0,blend_radius_m)
  movel([0.256303, -1.345181, -2.573748, -0.793461, 1.570796, 1.827100],accel_mss,speed_ms,0,blend_radius_m)
  movel([0.255412, -1.345809, -2.573331, -0.793249, 1.570796, 1.826209],accel_mss,speed_ms,0,blend_radius_m)
  movel([0.254724, -1.346319, -2.572992, -0.793078, 1.570796, 1.825520],accel_mss,speed_ms,0,blend_radius_m)
  movel([0.254047, -1.346846, -2.572641, -0.792902, 1.570796, 1.824843],accel_mss,speed_ms,0,blend_radius_m)
  movel([0.252379, -1.348218, -2.571726, -0.792445, 1.570796, 1.823175],accel_mss,speed_ms,0,blend_radius_m)
  movel([0.250748, -1.349634, -2.570780, -0.791975, 1.570796, 1.821544],accel_mss,speed_ms,0,blend_radius_m)
  movel([0.250109, -1.350216, -2.570389, -0.791783, 1.570796, 1.820906],accel_mss,speed_ms,0,blend_radius_m)
  movel([0.249486, -1.350814, -2.569988, -0.791586, 1.570796, 1.820283],accel_mss,speed_ms,0,blend_radius_m)
  movel([0.248861, -1.351441, -2.569568, -0.791380, 1.570796, 1.819657],accel_mss,speed_ms,0,blend_radius_m)
  movel([0.248252, -1.352078, -2.569139, -0.791172, 1.570796, 1.819048],accel_mss,speed_ms,0,blend_radius_m)
  movel([0.247658, -1.352723, -2.568705, -0.790961, 1.570796, 1.818454],accel_mss,speed_ms,0,blend_radius_m)
  movel([0.247081, -1.353376, -2.568265, -0.790748, 1.570796, 1.817877],accel_mss,speed_ms,0,blend_radius_m)
  movel([0.246522, -1.354036, -2.567819, -0.790534, 1.570796, 1.817318],accel_mss,speed_ms,0,blend_radius_m)
  movel([0.245984, -1.354698, -2.567372, -0.790320, 1.570796, 1.816781],accel_mss,speed_ms,0,blend_radius_m)
  movel([0.245466, -1.355366, -2.566919, -0.790104, 1.570796, 1.816263],accel_mss,speed_ms,0,blend_radius_m)
  movel([0.244966, -1.356040, -2.566463, -0.789886, 1.570796, 1.815763],accel_mss,speed_ms,0,blend_radius_m)
  movel([0.244487, -1.356719, -2.566002, -0.789668, 1.570796, 1.815283],accel_mss,speed_ms,0,blend_radius_m)
  movel([0.244025, -1.357403, -2.565537, -0.789449, 1.570796, 1.814821],accel_mss,speed_ms,0,blend_radius_m)
  movel([0.243592, -1.358077, -2.565078, -0.789234, 1.570796, 1.814388],accel_mss,speed_ms,0,blend_radius_m)
  movel([0.243180, -1.358754, -2.564616, -0.789018, 1.570796, 1.813976],accel_mss,speed_ms,0,blend_radius_m)
  movel([0.242791, -1.359434, -2.564153, -0.788803, 1.570796, 1.813587],accel_mss,speed_ms,0,blend_radius_m)
  movel([0.242421, -1.360114, -2.563688, -0.788587, 1.570796, 1.813217],accel_mss,speed_ms,0,blend_radius_m)
  movel([0.242071, -1.360799, -2.563219, -0.788371, 1.570796, 1.812867],accel_mss,speed_ms,0,blend_radius_m)
  movel([0.241755, -1.361462, -2.562765, -0.788162, 1.570796, 1.812551],accel_mss,speed_ms,0,blend_radius_m)
  movel([0.241459, -1.362128, -2.562307, -0.787953, 1.570796, 1.812256],accel_mss,speed_ms,0,blend_radius_m)
  movel([0.241191, -1.362792, -2.561852, -0.787746, 1.570796, 1.811987],accel_mss,speed_ms,0,blend_radius_m)
  movel([0.240944, -1.363453, -2.561396, -0.787539, 1.570796, 1.811740],accel_mss,speed_ms,0,blend_radius_m)
  movel([0.240721, -1.364112, -2.560942, -0.787334, 1.570796, 1.811517],accel_mss,speed_ms,0,blend_radius_m)
  movel([0.240451, -1.365015, -2.560320, -0.787055, 1.570796, 1.811247],accel_mss,speed_ms,0,blend_radius_m)
  movel([0.240217, -1.365913, -2.559699, -0.786777, 1.570796, 1.811013],accel_mss,speed_ms,0,blend_radius_m)
  movel([0.239938, -1.367112, -2.558868, -0.786409, 1.570796, 1.810734],accel_mss,speed_ms,0,blend_radius_m)
  movel([0.239680, -1.368307, -2.558038, -0.786044, 1.570796, 1.810476],accel_mss,speed_ms,0,blend_radius_m)
  movel([0.239448, -1.369472, -2.557228, -0.785690, 1.570796, 1.810244],accel_mss,speed_ms,0,blend_radius_m)
  movel([0.239237, -1.370627, -2.556422, -0.785341, 1.570796, 1.810033],accel_mss,speed_ms,0,blend_radius_m)
  movel([0.239129, -1.371375, -2.555899, -0.785115, 1.570796, 1.809925],accel_mss,speed_ms,0,blend_radius_m)
  movel([0.239064, -1.372107, -2.555386, -0.784896, 1.570796, 1.809860],accel_mss,speed_ms,0,blend_radius_m)
  movel([0.239040, -1.372671, -2.554991, -0.784727, 1.570796, 1.809837],accel_mss,speed_ms,0,blend_radius_m)
  movel([0.239038, -1.373226, -2.554601, -0.784561, 1.570796, 1.809834],accel_mss,speed_ms,0,blend_radius_m)
  movel([0.239055, -1.373774, -2.554216, -0.784398, 1.570796, 1.809852],accel_mss,speed_ms,0,blend_radius_m)
  movel([0.239094, -1.374314, -2.553837, -0.784238, 1.570796, 1.809890],accel_mss,speed_ms,0,blend_radius_m)
  movel([0.239153, -1.374844, -2.553464, -0.784081, 1.570796, 1.809949],accel_mss,speed_ms,0,blend_radius_m)
  movel([0.239230, -1.375366, -2.553096, -0.783927, 1.570796, 1.810026],accel_mss,speed_ms,0,blend_radius_m)
  movel([0.239326, -1.375877, -2.552735, -0.783777, 1.570796, 1.810122],accel_mss,speed_ms,0,blend_radius_m)
  movel([0.239469, -1.376486, -2.552305, -0.783598, 1.570796, 1.810266],accel_mss,speed_ms,0,blend_radius_m)
  movel([0.239636, -1.377085, -2.551881, -0.783422, 1.570796, 1.810432],accel_mss,speed_ms,0,blend_radius_m)
  movel([0.239830, -1.377667, -2.551470, -0.783252, 1.570796, 1.810626],accel_mss,speed_ms,0,blend_radius_m)
  movel([0.240045, -1.378236, -2.551066, -0.783087, 1.570796, 1.810841],accel_mss,speed_ms,0,blend_radius_m)
  movel([0.240284, -1.378789, -2.550674, -0.782926, 1.570796, 1.811081],accel_mss,speed_ms,0,blend_radius_m)
  movel([0.240546, -1.379327, -2.550292, -0.782770, 1.570796, 1.811342],accel_mss,speed_ms,0,blend_radius_m)
  movel([0.240841, -1.379866, -2.549908, -0.782614, 1.570796, 1.811637],accel_mss,speed_ms,0,blend_radius_m)
  movel([0.241158, -1.380389, -2.549536, -0.782464, 1.570796, 1.811955],accel_mss,speed_ms,0,blend_radius_m)
  movel([0.241499, -1.380894, -2.549177, -0.782319, 1.570796, 1.812295],accel_mss,speed_ms,0,blend_radius_m)
  movel([0.241860, -1.381384, -2.548827, -0.782178, 1.570796, 1.812657],accel_mss,speed_ms,0,blend_radius_m)
  movel([0.242243, -1.381854, -2.548491, -0.782044, 1.570796, 1.813039],accel_mss,speed_ms,0,blend_radius_m)
  movel([0.242648, -1.382308, -2.548167, -0.781914, 1.570796, 1.813444],accel_mss,speed_ms,0,blend_radius_m)
  movel([0.243080, -1.382749, -2.547851, -0.781788, 1.570796, 1.813877],accel_mss,speed_ms,0,blend_radius_m)
  movel([0.243531, -1.383173, -2.547548, -0.781668, 1.570796, 1.814327],accel_mss,speed_ms,0,blend_radius_m)
  movel([0.244002, -1.383579, -2.547257, -0.781553, 1.570796, 1.814798],accel_mss,speed_ms,0,blend_radius_m)
  movel([0.244493, -1.383965, -2.546980, -0.781443, 1.570796, 1.815290],accel_mss,speed_ms,0,blend_radius_m)
  movel([0.245003, -1.384334, -2.546716, -0.781339, 1.570796, 1.815799],accel_mss,speed_ms,0,blend_radius_m)
  movel([0.245528, -1.384683, -2.546465, -0.781241, 1.570796, 1.816325],accel_mss,speed_ms,0,blend_radius_m)
  movel([0.246115, -1.385035, -2.546212, -0.781142, 1.570796, 1.816911],accel_mss,speed_ms,0,blend_radius_m)
  movel([0.246714, -1.385368, -2.545973, -0.781048, 1.570796, 1.817511],accel_mss,speed_ms,0,blend_radius_m)
  movel([0.247335, -1.385679, -2.545749, -0.780961, 1.570796, 1.818132],accel_mss,speed_ms,0,blend_radius_m)
  movel([0.247973, -1.385969, -2.545540, -0.780880, 1.570796, 1.818769],accel_mss,speed_ms,0,blend_radius_m)
  movel([0.248627, -1.386238, -2.545347, -0.780804, 1.570796, 1.819423],accel_mss,speed_ms,0,blend_radius_m)
  movel([0.249299, -1.386484, -2.545170, -0.780736, 1.570796, 1.820095],accel_mss,speed_ms,0,blend_radius_m)
  movel([0.250013, -1.386719, -2.545000, -0.780670, 1.570796, 1.820810],accel_mss,speed_ms,0,blend_radius_m)
  movel([0.250744, -1.386937, -2.544843, -0.780609, 1.570796, 1.821540],accel_mss,speed_ms,0,blend_radius_m)
  movel([0.251487, -1.387134, -2.544701, -0.780555, 1.570796, 1.822283],accel_mss,speed_ms,0,blend_radius_m)
  movel([0.252244, -1.387308, -2.544575, -0.780506, 1.570796, 1.823041],accel_mss,speed_ms,0,blend_radius_m)
  movel([0.253013, -1.387464, -2.544462, -0.780463, 1.570796, 1.823810],accel_mss,speed_ms,0,blend_radius_m)
  movel([0.253794, -1.387601, -2.544363, -0.780425, 1.570796, 1.824591],accel_mss,speed_ms,0,blend_radius_m)
  movel([0.254605, -1.387719, -2.544278, -0.780392, 1.570796, 1.825401],accel_mss,speed_ms,0,blend_radius_m)
  movel([0.255429, -1.387815, -2.544209, -0.780365, 1.570796, 1.826225],accel_mss,speed_ms,0,blend_radius_m)
  movel([0.256261, -1.387893, -2.544152, -0.780344, 1.570796, 1.827058],accel_mss,speed_ms,0,blend_radius_m)
  movel([0.257105, -1.387950, -2.544111, -0.780328, 1.570796, 1.827901],accel_mss,speed_ms,0,blend_radius_m)
  movel([0.257958, -1.387985, -2.544086, -0.780318, 1.570796, 1.828755],accel_mss,speed_ms,0,blend_radius_m)
  movel([0.258821, -1.388002, -2.544073, -0.780313, 1.570796, 1.829617],accel_mss,speed_ms,0,blend_radius_m)
  movel([0.259693, -1.387996, -2.544078, -0.780315, 1.570796, 1.830489],accel_mss,speed_ms,0,blend_radius_m)
  movel([0.260575, -1.387970, -2.544097, -0.780322, 1.570796, 1.831371],accel_mss,speed_ms,0,blend_radius_m)
  movel([0.261462, -1.387925, -2.544129, -0.780335, 1.570796, 1.832259],accel_mss,speed_ms,0,blend_radius_m)
  movel([0.262358, -1.387858, -2.544178, -0.780353, 1.570796, 1.833154],accel_mss,speed_ms,0,blend_radius_m)
  movel([0.263262, -1.387770, -2.544241, -0.780378, 1.570796, 1.834059],accel_mss,speed_ms,0,blend_radius_m)
  movel([0.264172, -1.387663, -2.544319, -0.780407, 1.570796, 1.834968],accel_mss,speed_ms,0,blend_radius_m)
  movel([0.266174, -1.387406, -2.544504, -0.780479, 1.570796, 1.836970],accel_mss,speed_ms,0,blend_radius_m)
  movel([0.265950, -1.388175, -2.543948, -0.780265, 1.570796, 1.836746],accel_mss,speed_ms,0,blend_radius_m)
  movel([0.265726, -1.388944, -2.543392, -0.780053, 1.570796, 1.836522],accel_mss,speed_ms,0,blend_radius_m)
  movel([0.244685, -1.391802, -2.541316, -0.779271, 1.570796, 1.815481],accel_mss,speed_ms,0,blend_radius_m)
  movel([0.223610, -1.395032, -2.538956, -0.778401, 1.570796, 1.794406],accel_mss,speed_ms,0,blend_radius_m)
  movel([0.230335, -1.368198, -2.558114, -0.786077, 1.570796, 1.801132],accel_mss,speed_ms,0,blend_radius_m)
  movel([0.237492, -1.340228, -2.577017, -0.795144, 1.570796, 1.808288],accel_mss,speed_ms,0,blend_radius_m)
  movel([0.259913, -1.336512, -2.579449, -0.796428, 1.570796, 1.830709],accel_mss,speed_ms,0,blend_radius_m)
  movel([0.282293, -1.333219, -2.581588, -0.797582, 1.570796, 1.853089],accel_mss,speed_ms,0,blend_radius_m)
  speed_ms = 0.003
  movel([0.282293, -1.336450, -2.583168, -0.792771, 1.570796, 1.853089],accel_mss,speed_ms,0,blend_radius_m)
  speed_ms = 0.007
  movel([0.281918, -1.337684, -2.582364, -0.792340, 1.570796, 1.852714],accel_mss,speed_ms,0,blend_radius_m)
  movel([0.281544, -1.338916, -2.581560, -0.791913, 1.570796, 1.852341],accel_mss,speed_ms,0,blend_radius_m)
  movel([0.278441, -1.339413, -2.581235, -0.791741, 1.570796, 1.849238],accel_mss,speed_ms,0,blend_radius_m)
  movel([0.276251, -1.339793, -2.580986, -0.791610, 1.570796, 1.847047],accel_mss,speed_ms,0,blend_radius_m)
  movel([0.275394, -1.339962, -2.580875, -0.791551, 1.570796, 1.846190],accel_mss,speed_ms,0,blend_radius_m)
  movel([0.274530, -1.340156, -2.580749, -0.791485, 1.570796, 1.845326],accel_mss,speed_ms,0,blend_radius_m)
  movel([0.273708, -1.340359, -2.580615, -0.791415, 1.570796, 1.844505],accel_mss,speed_ms,0,blend_radius_m)
  movel([0.272883, -1.340584, -2.580467, -0.791337, 1.570796, 1.843679],accel_mss,speed_ms,0,blend_radius_m)
  movel([0.270940, -1.341174, -2.580081, -0.791135, 1.570796, 1.841736],accel_mss,speed_ms,0,blend_radius_m)
  movel([0.269926, -1.341509, -2.579860, -0.791020, 1.570796, 1.840722],accel_mss,speed_ms,0,blend_radius_m)
  movel([0.268912, -1.341870, -2.579623, -0.790896, 1.570796, 1.839708],accel_mss,speed_ms,0,blend_radius_m)
  movel([0.267897, -1.342252, -2.579371, -0.790765, 1.570796, 1.838694],accel_mss,speed_ms,0,blend_radius_m)
  movel([0.266884, -1.342657, -2.579105, -0.790627, 1.570796, 1.837680],accel_mss,speed_ms,0,blend_radius_m)
  movel([0.265880, -1.343082, -2.578825, -0.790482, 1.570796, 1.836676],accel_mss,speed_ms,0,blend_radius_m)
  movel([0.264877, -1.343529, -2.578530, -0.790330, 1.570796, 1.835673],accel_mss,speed_ms,0,blend_radius_m)
  movel([0.263878, -1.343999, -2.578220, -0.790171, 1.570796, 1.834675],accel_mss,speed_ms,0,blend_radius_m)
  movel([0.262881, -1.344489, -2.577896, -0.790005, 1.570796, 1.833678],accel_mss,speed_ms,0,blend_radius_m)
  movel([0.261910, -1.344993, -2.577562, -0.789834, 1.570796, 1.832706],accel_mss,speed_ms,0,blend_radius_m)
  movel([0.260943, -1.345517, -2.577215, -0.789657, 1.570796, 1.831739],accel_mss,speed_ms,0,blend_radius_m)
  movel([0.259983, -1.346061, -2.576855, -0.789474, 1.570796, 1.830780],accel_mss,speed_ms,0,blend_radius_m)
  movel([0.259028, -1.346626, -2.576479, -0.789284, 1.570796, 1.829824],accel_mss,speed_ms,0,blend_radius_m)
  movel([0.258111, -1.347192, -2.576103, -0.789094, 1.570796, 1.828907],accel_mss,speed_ms,0,blend_radius_m)
  movel([0.257201, -1.347780, -2.575712, -0.788897, 1.570796, 1.827997],accel_mss,speed_ms,0,blend_radius_m)
  movel([0.256303, -1.348386, -2.575308, -0.788695, 1.570796, 1.827100],accel_mss,speed_ms,0,blend_radius_m)
  movel([0.255412, -1.349012, -2.574890, -0.788486, 1.570796, 1.826209],accel_mss,speed_ms,0,blend_radius_m)
  movel([0.254724, -1.349521, -2.574551, -0.788317, 1.570796, 1.825520],accel_mss,speed_ms,0,blend_radius_m)
  movel([0.254047, -1.350047, -2.574199, -0.788143, 1.570796, 1.824843],accel_mss,speed_ms,0,blend_radius_m)
  movel([0.252379, -1.351416, -2.573282, -0.787691, 1.570796, 1.823175],accel_mss,speed_ms,0,blend_radius_m)
  movel([0.250748, -1.352829, -2.572333, -0.787227, 1.570796, 1.821544],accel_mss,speed_ms,0,blend_radius_m)
  movel([0.250109, -1.353410, -2.571942, -0.787037, 1.570796, 1.820906],accel_mss,speed_ms,0,blend_radius_m)
  movel([0.249486, -1.354006, -2.571540, -0.786843, 1.570796, 1.820283],accel_mss,speed_ms,0,blend_radius_m)
  movel([0.248861, -1.354631, -2.571118, -0.786639, 1.570796, 1.819657],accel_mss,speed_ms,0,blend_radius_m)
  movel([0.248252, -1.355267, -2.570689, -0.786433, 1.570796, 1.819048],accel_mss,speed_ms,0,blend_radius_m)
  movel([0.247658, -1.355910, -2.570253, -0.786225, 1.570796, 1.818454],accel_mss,speed_ms,0,blend_radius_m)
  movel([0.247081, -1.356562, -2.569812, -0.786015, 1.570796, 1.817877],accel_mss,speed_ms,0,blend_radius_m)
  movel([0.246522, -1.357221, -2.569365, -0.785803, 1.570796, 1.817318],accel_mss,speed_ms,0,blend_radius_m)
  movel([0.245984, -1.357881, -2.568917, -0.785591, 1.570796, 1.816781],accel_mss,speed_ms,0,blend_radius_m)
  movel([0.245466, -1.358548, -2.568464, -0.785378, 1.570796, 1.816263],accel_mss,speed_ms,0,blend_radius_m)
  movel([0.244966, -1.359220, -2.568006, -0.785163, 1.570796, 1.815763],accel_mss,speed_ms,0,blend_radius_m)
  movel([0.244487, -1.359897, -2.567544, -0.784948, 1.570796, 1.815283],accel_mss,speed_ms,0,blend_radius_m)
  movel([0.244025, -1.360580, -2.567078, -0.784732, 1.570796, 1.814821],accel_mss,speed_ms,0,blend_radius_m)
  movel([0.243592, -1.361253, -2.566618, -0.784519, 1.570796, 1.814388],accel_mss,speed_ms,0,blend_radius_m)
  movel([0.243180, -1.361928, -2.566155, -0.784306, 1.570796, 1.813976],accel_mss,speed_ms,0,blend_radius_m)
  movel([0.242791, -1.362606, -2.565690, -0.784093, 1.570796, 1.813587],accel_mss,speed_ms,0,blend_radius_m)
  movel([0.242421, -1.363284, -2.565224, -0.783880, 1.570796, 1.813217],accel_mss,speed_ms,0,blend_radius_m)
  movel([0.242071, -1.363968, -2.564755, -0.783667, 1.570796, 1.812867],accel_mss,speed_ms,0,blend_radius_m)
  movel([0.241755, -1.364630, -2.564299, -0.783461, 1.570796, 1.812551],accel_mss,speed_ms,0,blend_radius_m)
  movel([0.241459, -1.365294, -2.563841, -0.783254, 1.570796, 1.812256],accel_mss,speed_ms,0,blend_radius_m)
  movel([0.241191, -1.365956, -2.563384, -0.783049, 1.570796, 1.811987],accel_mss,speed_ms,0,blend_radius_m)
  movel([0.240944, -1.366616, -2.562927, -0.782846, 1.570796, 1.811740],accel_mss,speed_ms,0,blend_radius_m)
  movel([0.240721, -1.367274, -2.562472, -0.782643, 1.570796, 1.811517],accel_mss,speed_ms,0,blend_radius_m)
  movel([0.240451, -1.368174, -2.561848, -0.782367, 1.570796, 1.811247],accel_mss,speed_ms,0,blend_radius_m)
  movel([0.240217, -1.369070, -2.561226, -0.782093, 1.570796, 1.811013],accel_mss,speed_ms,0,blend_radius_m)
  movel([0.239938, -1.370267, -2.560393, -0.781730, 1.570796, 1.810734],accel_mss,speed_ms,0,blend_radius_m)
  movel([0.239680, -1.371458, -2.559561, -0.781369, 1.570796, 1.810476],accel_mss,speed_ms,0,blend_radius_m)
  movel([0.239448, -1.372620, -2.558749, -0.781020, 1.570796, 1.810244],accel_mss,speed_ms,0,blend_radius_m)
  movel([0.239237, -1.373773, -2.557941, -0.780675, 1.570796, 1.810033],accel_mss,speed_ms,0,blend_radius_m)
  movel([0.239129, -1.374519, -2.557417, -0.780453, 1.570796, 1.809925],accel_mss,speed_ms,0,blend_radius_m)
  movel([0.239064, -1.375249, -2.556903, -0.780236, 1.570796, 1.809860],accel_mss,speed_ms,0,blend_radius_m)
  movel([0.239040, -1.375811, -2.556507, -0.780070, 1.570796, 1.809837],accel_mss,speed_ms,0,blend_radius_m)
  movel([0.239038, -1.376366, -2.556117, -0.779907, 1.570796, 1.809834],accel_mss,speed_ms,0,blend_radius_m)
  movel([0.239055, -1.376912, -2.555731, -0.779746, 1.570796, 1.809852],accel_mss,speed_ms,0,blend_radius_m)
  movel([0.239094, -1.377451, -2.555350, -0.779588, 1.570796, 1.809890],accel_mss,speed_ms,0,blend_radius_m)
  movel([0.239153, -1.377979, -2.554976, -0.779433, 1.570796, 1.809949],accel_mss,speed_ms,0,blend_radius_m)
  movel([0.239230, -1.378501, -2.554607, -0.779281, 1.570796, 1.810026],accel_mss,speed_ms,0,blend_radius_m)
  movel([0.239326, -1.379010, -2.554246, -0.779133, 1.570796, 1.810122],accel_mss,speed_ms,0,blend_radius_m)
  movel([0.239469, -1.379618, -2.553815, -0.778956, 1.570796, 1.810266],accel_mss,speed_ms,0,blend_radius_m)
  movel([0.239636, -1.380216, -2.553390, -0.778783, 1.570796, 1.810432],accel_mss,speed_ms,0,blend_radius_m)
  movel([0.239830, -1.380796, -2.552978, -0.778615, 1.570796, 1.810626],accel_mss,speed_ms,0,blend_radius_m)
  movel([0.240045, -1.381364, -2.552573, -0.778452, 1.570796, 1.810841],accel_mss,speed_ms,0,blend_radius_m)
  movel([0.240284, -1.381915, -2.552180, -0.778294, 1.570796, 1.811081],accel_mss,speed_ms,0,blend_radius_m)
  movel([0.240546, -1.382452, -2.551797, -0.778140, 1.570796, 1.811342],accel_mss,speed_ms,0,blend_radius_m)
  movel([0.240841, -1.382990, -2.551413, -0.777986, 1.570796, 1.811637],accel_mss,speed_ms,0,blend_radius_m)
  movel([0.241158, -1.383512, -2.551040, -0.777838, 1.570796, 1.811955],accel_mss,speed_ms,0,blend_radius_m)
  movel([0.241499, -1.384015, -2.550680, -0.777695, 1.570796, 1.812295],accel_mss,speed_ms,0,blend_radius_m)
  movel([0.241860, -1.384504, -2.550329, -0.777556, 1.570796, 1.812657],accel_mss,speed_ms,0,blend_radius_m)
  movel([0.242243, -1.384973, -2.549993, -0.777423, 1.570796, 1.813039],accel_mss,speed_ms,0,blend_radius_m)
  movel([0.242648, -1.385426, -2.549668, -0.777296, 1.570796, 1.813444],accel_mss,speed_ms,0,blend_radius_m)
  movel([0.243080, -1.385866, -2.549351, -0.777172, 1.570796, 1.813877],accel_mss,speed_ms,0,blend_radius_m)
  movel([0.243531, -1.386288, -2.549047, -0.777053, 1.570796, 1.814327],accel_mss,speed_ms,0,blend_radius_m)
  movel([0.244002, -1.386693, -2.548756, -0.776940, 1.570796, 1.814798],accel_mss,speed_ms,0,blend_radius_m)
  movel([0.244493, -1.387079, -2.548479, -0.776832, 1.570796, 1.815290],accel_mss,speed_ms,0,blend_radius_m)
  movel([0.245003, -1.387446, -2.548213, -0.776729, 1.570796, 1.815799],accel_mss,speed_ms,0,blend_radius_m)
  movel([0.245528, -1.387795, -2.547962, -0.776632, 1.570796, 1.816325],accel_mss,speed_ms,0,blend_radius_m)
  movel([0.246115, -1.388146, -2.547709, -0.776534, 1.570796, 1.816911],accel_mss,speed_ms,0,blend_radius_m)
  movel([0.246714, -1.388478, -2.547469, -0.776442, 1.570796, 1.817511],accel_mss,speed_ms,0,blend_radius_m)
  movel([0.247335, -1.388788, -2.547245, -0.776356, 1.570796, 1.818132],accel_mss,speed_ms,0,blend_radius_m)
  movel([0.247973, -1.389077, -2.547035, -0.776276, 1.570796, 1.818769],accel_mss,speed_ms,0,blend_radius_m)
  movel([0.248627, -1.389346, -2.546841, -0.776202, 1.570796, 1.819423],accel_mss,speed_ms,0,blend_radius_m)
  movel([0.249299, -1.389591, -2.546664, -0.776134, 1.570796, 1.820095],accel_mss,speed_ms,0,blend_radius_m)
  movel([0.250013, -1.389826, -2.546493, -0.776069, 1.570796, 1.820810],accel_mss,speed_ms,0,blend_radius_m)
  movel([0.250744, -1.390043, -2.546336, -0.776010, 1.570796, 1.821540],accel_mss,speed_ms,0,blend_radius_m)
  movel([0.251487, -1.390239, -2.546194, -0.775956, 1.570796, 1.822283],accel_mss,speed_ms,0,blend_radius_m)
  movel([0.252244, -1.390413, -2.546068, -0.775908, 1.570796, 1.823041],accel_mss,speed_ms,0,blend_radius_m)
  movel([0.253013, -1.390569, -2.545954, -0.775865, 1.570796, 1.823810],accel_mss,speed_ms,0,blend_radius_m)
  movel([0.253794, -1.390705, -2.545856, -0.775828, 1.570796, 1.824591],accel_mss,speed_ms,0,blend_radius_m)
  movel([0.254605, -1.390823, -2.545770, -0.775795, 1.570796, 1.825401],accel_mss,speed_ms,0,blend_radius_m)
  movel([0.255429, -1.390919, -2.545701, -0.775769, 1.570796, 1.826225],accel_mss,speed_ms,0,blend_radius_m)
  movel([0.256261, -1.390997, -2.545644, -0.775748, 1.570796, 1.827058],accel_mss,speed_ms,0,blend_radius_m)
  movel([0.257105, -1.391054, -2.545603, -0.775732, 1.570796, 1.827901],accel_mss,speed_ms,0,blend_radius_m)
  movel([0.257958, -1.391088, -2.545578, -0.775723, 1.570796, 1.828755],accel_mss,speed_ms,0,blend_radius_m)
  movel([0.258821, -1.391106, -2.545565, -0.775718, 1.570796, 1.829617],accel_mss,speed_ms,0,blend_radius_m)
  movel([0.259693, -1.391099, -2.545570, -0.775720, 1.570796, 1.830489],accel_mss,speed_ms,0,blend_radius_m)
  movel([0.260575, -1.391073, -2.545589, -0.775727, 1.570796, 1.831371],accel_mss,speed_ms,0,blend_radius_m)
  movel([0.261462, -1.391028, -2.545621, -0.775739, 1.570796, 1.832259],accel_mss,speed_ms,0,blend_radius_m)
  movel([0.262358, -1.390962, -2.545669, -0.775757, 1.570796, 1.833154],accel_mss,speed_ms,0,blend_radius_m)
  movel([0.263262, -1.390874, -2.545733, -0.775782, 1.570796, 1.834059],accel_mss,speed_ms,0,blend_radius_m)
  movel([0.264172, -1.390767, -2.545811, -0.775811, 1.570796, 1.834968],accel_mss,speed_ms,0,blend_radius_m)
  movel([0.266174, -1.390511, -2.545997, -0.775881, 1.570796, 1.836970],accel_mss,speed_ms,0,blend_radius_m)
  movel([0.265950, -1.391279, -2.545440, -0.775671, 1.570796, 1.836746],accel_mss,speed_ms,0,blend_radius_m)
  movel([0.265726, -1.392045, -2.544882, -0.775462, 1.570796, 1.836522],accel_mss,speed_ms,0,blend_radius_m)
  movel([0.244685, -1.394897, -2.542801, -0.774691, 1.570796, 1.815481],accel_mss,speed_ms,0,blend_radius_m)
  movel([0.223610, -1.398118, -2.540436, -0.773834, 1.570796, 1.794406],accel_mss,speed_ms,0,blend_radius_m)
  movel([0.230335, -1.371349, -2.559638, -0.781402, 1.570796, 1.801132],accel_mss,speed_ms,0,blend_radius_m)
  movel([0.237492, -1.343444, -2.578586, -0.790359, 1.570796, 1.808288],accel_mss,speed_ms,0,blend_radius_m)
  movel([0.259913, -1.339736, -2.581023, -0.791629, 1.570796, 1.830709],accel_mss,speed_ms,0,blend_radius_m)
  movel([0.282293, -1.336450, -2.583168, -0.792771, 1.570796, 1.853089],accel_mss,speed_ms,0,blend_radius_m)
  speed_ms = 0.003
  movel([0.282293, -1.323668, -2.576799, -0.811922, 1.570796, 1.853089],accel_mss,speed_ms,0,blend_radius_m)
  speed_ms = 0.01
  movel([0.282293, -1.299239, -2.563684, -0.849465, 1.570796, 1.853089],accel_mss,speed_ms,0,blend_radius_m)
  movel([0.280179, -1.305078, -2.560060, -0.847250, 1.570796, 1.850975],accel_mss,speed_ms,0,blend_radius_m)
  movel([0.280179, -1.329425, -2.573101, -0.809863, 1.570796, 1.850975],accel_mss,speed_ms,0,blend_radius_m)
  speed_ms = 0.003
  movel([0.280179, -1.338941, -2.577862, -0.795587, 1.570796, 1.850975],accel_mss,speed_ms,0,blend_radius_m)
  speed_ms = 0.007
  movel([0.280440, -1.338973, -2.577841, -0.795576, 1.570796, 1.851236],accel_mss,speed_ms,0,blend_radius_m)
  movel([0.273536, -1.361801, -2.562532, -0.788056, 1.570796, 1.844333],accel_mss,speed_ms,0,blend_radius_m)
  movel([0.270969, -1.370377, -2.556596, -0.785416, 1.570796, 1.841766],accel_mss,speed_ms,0,blend_radius_m)
  movel([0.268811, -1.377594, -2.551521, -0.783274, 1.570796, 1.839607],accel_mss,speed_ms,0,blend_radius_m)
  movel([0.266912, -1.383952, -2.546990, -0.781447, 1.570796, 1.837709],accel_mss,speed_ms,0,blend_radius_m)
  movel([0.266850, -1.384141, -2.546855, -0.781394, 1.570796, 1.837647],accel_mss,speed_ms,0,blend_radius_m)
  movel([0.266777, -1.384331, -2.546718, -0.781340, 1.570796, 1.837573],accel_mss,speed_ms,0,blend_radius_m)
  movel([0.266578, -1.384809, -2.546375, -0.781205, 1.570796, 1.837374],accel_mss,speed_ms,0,blend_radius_m)
  movel([0.264610, -1.385063, -2.546192, -0.781134, 1.570796, 1.835406],accel_mss,speed_ms,0,blend_radius_m)
  movel([0.263843, -1.385154, -2.546127, -0.781108, 1.570796, 1.834640],accel_mss,speed_ms,0,blend_radius_m)
  movel([0.263083, -1.385230, -2.546072, -0.781087, 1.570796, 1.833879],accel_mss,speed_ms,0,blend_radius_m)
  movel([0.262327, -1.385291, -2.546028, -0.781070, 1.570796, 1.833124],accel_mss,speed_ms,0,blend_radius_m)
  movel([0.261578, -1.385337, -2.545995, -0.781057, 1.570796, 1.832375],accel_mss,speed_ms,0,blend_radius_m)
  movel([0.260834, -1.385366, -2.545974, -0.781049, 1.570796, 1.831630],accel_mss,speed_ms,0,blend_radius_m)
  movel([0.260096, -1.385382, -2.545963, -0.781044, 1.570796, 1.830892],accel_mss,speed_ms,0,blend_radius_m)
  movel([0.259365, -1.385380, -2.545964, -0.781045, 1.570796, 1.830161],accel_mss,speed_ms,0,blend_radius_m)
  movel([0.258640, -1.385363, -2.545976, -0.781049, 1.570796, 1.829436],accel_mss,speed_ms,0,blend_radius_m)
  movel([0.257923, -1.385329, -2.546001, -0.781059, 1.570796, 1.828719],accel_mss,speed_ms,0,blend_radius_m)
  movel([0.257213, -1.385281, -2.546035, -0.781072, 1.570796, 1.828010],accel_mss,speed_ms,0,blend_radius_m)
  movel([0.256522, -1.385217, -2.546081, -0.781091, 1.570796, 1.827318],accel_mss,speed_ms,0,blend_radius_m)
  movel([0.255839, -1.385139, -2.546137, -0.781112, 1.570796, 1.826635],accel_mss,speed_ms,0,blend_radius_m)
  movel([0.255166, -1.385044, -2.546206, -0.781139, 1.570796, 1.825962],accel_mss,speed_ms,0,blend_radius_m)
  movel([0.254501, -1.384930, -2.546288, -0.781171, 1.570796, 1.825298],accel_mss,speed_ms,0,blend_radius_m)
  movel([0.253845, -1.384803, -2.546379, -0.781207, 1.570796, 1.824641],accel_mss,speed_ms,0,blend_radius_m)
  movel([0.253200, -1.384661, -2.546481, -0.781247, 1.570796, 1.823996],accel_mss,speed_ms,0,blend_radius_m)
  movel([0.252563, -1.384502, -2.546595, -0.781292, 1.570796, 1.823360],accel_mss,speed_ms,0,blend_radius_m)
  movel([0.251938, -1.384328, -2.546720, -0.781341, 1.570796, 1.822734],accel_mss,speed_ms,0,blend_radius_m)
  movel([0.251323, -1.384138, -2.546857, -0.781395, 1.570796, 1.822119],accel_mss,speed_ms,0,blend_radius_m)
  movel([0.250721, -1.383931, -2.547005, -0.781453, 1.570796, 1.821518],accel_mss,speed_ms,0,blend_radius_m)
  movel([0.250151, -1.383718, -2.547158, -0.781513, 1.570796, 1.820947],accel_mss,speed_ms,0,blend_radius_m)
  movel([0.249594, -1.383489, -2.547322, -0.781578, 1.570796, 1.820390],accel_mss,speed_ms,0,blend_radius_m)
  movel([0.249050, -1.383245, -2.547497, -0.781647, 1.570796, 1.819846],accel_mss,speed_ms,0,blend_radius_m)
  movel([0.248516, -1.382985, -2.547683, -0.781721, 1.570796, 1.819312],accel_mss,speed_ms,0,blend_radius_m)
  movel([0.247995, -1.382711, -2.547879, -0.781799, 1.570796, 1.818792],accel_mss,speed_ms,0,blend_radius_m)
  movel([0.247488, -1.382420, -2.548087, -0.781882, 1.570796, 1.818284],accel_mss,speed_ms,0,blend_radius_m)
  movel([0.246994, -1.382117, -2.548303, -0.781968, 1.570796, 1.817791],accel_mss,speed_ms,0,blend_radius_m)
  movel([0.246515, -1.381797, -2.548532, -0.782060, 1.570796, 1.817311],accel_mss,speed_ms,0,blend_radius_m)
  movel([0.246047, -1.381463, -2.548771, -0.782155, 1.570796, 1.816844],accel_mss,speed_ms,0,blend_radius_m)
  movel([0.245597, -1.381116, -2.549018, -0.782255, 1.570796, 1.816393],accel_mss,speed_ms,0,blend_radius_m)
  movel([0.245219, -1.380802, -2.549242, -0.782345, 1.570796, 1.816016],accel_mss,speed_ms,0,blend_radius_m)
  movel([0.244858, -1.380478, -2.549473, -0.782438, 1.570796, 1.815654],accel_mss,speed_ms,0,blend_radius_m)
  movel([0.244510, -1.380139, -2.549714, -0.782536, 1.570796, 1.815306],accel_mss,speed_ms,0,blend_radius_m)
  movel([0.244175, -1.379789, -2.549963, -0.782637, 1.570796, 1.814972],accel_mss,speed_ms,0,blend_radius_m)
  movel([0.243853, -1.379427, -2.550220, -0.782741, 1.570796, 1.814649],accel_mss,speed_ms,0,blend_radius_m)
  movel([0.243548, -1.379052, -2.550487, -0.782850, 1.570796, 1.814344],accel_mss,speed_ms,0,blend_radius_m)
  movel([0.243259, -1.378664, -2.550763, -0.782962, 1.570796, 1.814056],accel_mss,speed_ms,0,blend_radius_m)
  movel([0.242982, -1.378267, -2.551044, -0.783078, 1.570796, 1.813778],accel_mss,speed_ms,0,blend_radius_m)
  movel([0.242723, -1.377855, -2.551337, -0.783198, 1.570796, 1.813519],accel_mss,speed_ms,0,blend_radius_m)
  movel([0.242476, -1.377434, -2.551635, -0.783320, 1.570796, 1.813273],accel_mss,speed_ms,0,blend_radius_m)
  movel([0.242247, -1.377002, -2.551941, -0.783447, 1.570796, 1.813043],accel_mss,speed_ms,0,blend_radius_m)
  movel([0.242044, -1.376578, -2.552240, -0.783571, 1.570796, 1.812841],accel_mss,speed_ms,0,blend_radius_m)
  movel([0.241857, -1.376141, -2.552549, -0.783699, 1.570796, 1.812653],accel_mss,speed_ms,0,blend_radius_m)
  movel([0.241688, -1.375695, -2.552864, -0.783830, 1.570796, 1.812484],accel_mss,speed_ms,0,blend_radius_m)
  movel([0.241534, -1.375240, -2.553185, -0.783964, 1.570796, 1.812331],accel_mss,speed_ms,0,blend_radius_m)
  movel([0.241400, -1.374773, -2.553514, -0.784102, 1.570796, 1.812197],accel_mss,speed_ms,0,blend_radius_m)
  movel([0.241282, -1.374297, -2.553849, -0.784243, 1.570796, 1.812078],accel_mss,speed_ms,0,blend_radius_m)
  movel([0.241179, -1.373814, -2.554189, -0.784387, 1.570796, 1.811976],accel_mss,speed_ms,0,blend_radius_m)
  movel([0.241096, -1.373319, -2.554536, -0.784534, 1.570796, 1.811892],accel_mss,speed_ms,0,blend_radius_m)
  movel([0.241030, -1.372817, -2.554889, -0.784684, 1.570796, 1.811827],accel_mss,speed_ms,0,blend_radius_m)
  movel([0.240983, -1.372307, -2.555246, -0.784836, 1.570796, 1.811779],accel_mss,speed_ms,0,blend_radius_m)
  movel([0.240954, -1.371796, -2.555604, -0.784989, 1.570796, 1.811750],accel_mss,speed_ms,0,blend_radius_m)
  movel([0.240943, -1.371277, -2.555967, -0.785145, 1.570796, 1.811739],accel_mss,speed_ms,0,blend_radius_m)
  movel([0.240950, -1.370752, -2.556335, -0.785303, 1.570796, 1.811746],accel_mss,speed_ms,0,blend_radius_m)
  movel([0.240977, -1.370218, -2.556707, -0.785464, 1.570796, 1.811774],accel_mss,speed_ms,0,blend_radius_m)
  movel([0.241023, -1.369679, -2.557083, -0.785627, 1.570796, 1.811819],accel_mss,speed_ms,0,blend_radius_m)
  movel([0.241086, -1.369134, -2.557463, -0.785792, 1.570796, 1.811882],accel_mss,speed_ms,0,blend_radius_m)
  movel([0.241165, -1.368587, -2.557844, -0.785959, 1.570796, 1.811962],accel_mss,speed_ms,0,blend_radius_m)
  movel([0.241266, -1.368031, -2.558230, -0.786128, 1.570796, 1.812062],accel_mss,speed_ms,0,blend_radius_m)
  movel([0.241384, -1.367472, -2.558618, -0.786299, 1.570796, 1.812180],accel_mss,speed_ms,0,blend_radius_m)
  movel([0.241521, -1.366910, -2.559008, -0.786471, 1.570796, 1.812317],accel_mss,speed_ms,0,blend_radius_m)
  movel([0.241675, -1.366344, -2.559400, -0.786644, 1.570796, 1.812471],accel_mss,speed_ms,0,blend_radius_m)
  movel([0.241849, -1.365775, -2.559794, -0.786820, 1.570796, 1.812645],accel_mss,speed_ms,0,blend_radius_m)
  movel([0.242040, -1.365205, -2.560188, -0.786996, 1.570796, 1.812836],accel_mss,speed_ms,0,blend_radius_m)
  movel([0.242247, -1.364635, -2.560582, -0.787172, 1.570796, 1.813043],accel_mss,speed_ms,0,blend_radius_m)
  movel([0.242474, -1.364060, -2.560978, -0.787351, 1.570796, 1.813270],accel_mss,speed_ms,0,blend_radius_m)
  movel([0.242718, -1.363484, -2.561375, -0.787530, 1.570796, 1.813514],accel_mss,speed_ms,0,blend_radius_m)
  movel([0.242978, -1.362910, -2.561770, -0.787709, 1.570796, 1.813774],accel_mss,speed_ms,0,blend_radius_m)
  movel([0.243257, -1.362335, -2.562166, -0.787889, 1.570796, 1.814053],accel_mss,speed_ms,0,blend_radius_m)
  movel([0.243552, -1.361761, -2.562560, -0.788069, 1.570796, 1.814348],accel_mss,speed_ms,0,blend_radius_m)
  movel([0.243864, -1.361188, -2.562953, -0.788249, 1.570796, 1.814660],accel_mss,speed_ms,0,blend_radius_m)
  movel([0.244196, -1.360609, -2.563349, -0.788431, 1.570796, 1.814992],accel_mss,speed_ms,0,blend_radius_m)
  movel([0.244544, -1.360034, -2.563743, -0.788613, 1.570796, 1.815340],accel_mss,speed_ms,0,blend_radius_m)
  movel([0.244905, -1.359463, -2.564133, -0.788793, 1.570796, 1.815701],accel_mss,speed_ms,0,blend_radius_m)
  movel([0.245284, -1.358892, -2.564522, -0.788974, 1.570796, 1.816081],accel_mss,speed_ms,0,blend_radius_m)
  movel([0.245678, -1.358324, -2.564910, -0.789155, 1.570796, 1.816475],accel_mss,speed_ms,0,blend_radius_m)
  movel([0.246085, -1.357762, -2.565293, -0.789334, 1.570796, 1.816881],accel_mss,speed_ms,0,blend_radius_m)
  movel([0.246509, -1.357205, -2.565671, -0.789512, 1.570796, 1.817305],accel_mss,speed_ms,0,blend_radius_m)
  movel([0.246944, -1.356651, -2.566048, -0.789690, 1.570796, 1.817741],accel_mss,speed_ms,0,blend_radius_m)
  movel([0.247394, -1.356105, -2.566418, -0.789865, 1.570796, 1.818191],accel_mss,speed_ms,0,blend_radius_m)
  movel([0.247858, -1.355563, -2.566786, -0.790040, 1.570796, 1.818654],accel_mss,speed_ms,0,blend_radius_m)
  movel([0.248368, -1.354989, -2.567174, -0.790225, 1.570796, 1.819164],accel_mss,speed_ms,0,blend_radius_m)
  movel([0.248888, -1.354425, -2.567556, -0.790408, 1.570796, 1.819684],accel_mss,speed_ms,0,blend_radius_m)
  movel([0.249421, -1.353867, -2.567934, -0.790589, 1.570796, 1.820217],accel_mss,speed_ms,0,blend_radius_m)
  movel([0.249964, -1.353315, -2.568306, -0.790768, 1.570796, 1.820760],accel_mss,speed_ms,0,blend_radius_m)
  movel([0.250520, -1.352771, -2.568673, -0.790946, 1.570796, 1.821316],accel_mss,speed_ms,0,blend_radius_m)
  movel([0.251085, -1.352237, -2.569032, -0.791120, 1.570796, 1.821881],accel_mss,speed_ms,0,blend_radius_m)
  movel([0.251663, -1.351708, -2.569388, -0.791293, 1.570796, 1.822460],accel_mss,speed_ms,0,blend_radius_m)
  movel([0.252248, -1.351192, -2.569735, -0.791462, 1.570796, 1.823045],accel_mss,speed_ms,0,blend_radius_m)
  movel([0.252844, -1.350682, -2.570077, -0.791630, 1.570796, 1.823640],accel_mss,speed_ms,0,blend_radius_m)
  movel([0.253467, -1.350170, -2.570421, -0.791798, 1.570796, 1.824263],accel_mss,speed_ms,0,blend_radius_m)
  movel([0.254097, -1.349665, -2.570759, -0.791965, 1.570796, 1.824893],accel_mss,speed_ms,0,blend_radius_m)
  movel([0.254735, -1.349171, -2.571090, -0.792129, 1.570796, 1.825531],accel_mss,speed_ms,0,blend_radius_m)
  movel([0.255380, -1.348686, -2.571414, -0.792289, 1.570796, 1.826176],accel_mss,speed_ms,0,blend_radius_m)
  movel([0.256033, -1.348213, -2.571730, -0.792446, 1.570796, 1.826830],accel_mss,speed_ms,0,blend_radius_m)
  movel([0.256692, -1.347751, -2.572038, -0.792600, 1.570796, 1.827488],accel_mss,speed_ms,0,blend_radius_m)
  movel([0.257360, -1.347298, -2.572340, -0.792751, 1.570796, 1.828157],accel_mss,speed_ms,0,blend_radius_m)
  movel([0.258033, -1.346857, -2.572633, -0.792898, 1.570796, 1.828829],accel_mss,speed_ms,0,blend_radius_m)
  movel([0.258710, -1.346428, -2.572919, -0.793042, 1.570796, 1.829506],accel_mss,speed_ms,0,blend_radius_m)
  movel([0.259422, -1.345993, -2.573209, -0.793188, 1.570796, 1.830218],accel_mss,speed_ms,0,blend_radius_m)
  movel([0.260138, -1.345568, -2.573490, -0.793330, 1.570796, 1.830935],accel_mss,speed_ms,0,blend_radius_m)
  movel([0.260861, -1.345159, -2.573762, -0.793468, 1.570796, 1.831657],accel_mss,speed_ms,0,blend_radius_m)
  movel([0.261586, -1.344760, -2.574027, -0.793602, 1.570796, 1.832382],accel_mss,speed_ms,0,blend_radius_m)
  movel([0.262317, -1.344374, -2.574282, -0.793732, 1.570796, 1.833113],accel_mss,speed_ms,0,blend_radius_m)
  movel([0.263049, -1.344002, -2.574529, -0.793858, 1.570796, 1.833845],accel_mss,speed_ms,0,blend_radius_m)
  movel([0.263783, -1.343642, -2.574767, -0.793980, 1.570796, 1.834579],accel_mss,speed_ms,0,blend_radius_m)
  movel([0.264523, -1.343296, -2.574996, -0.794097, 1.570796, 1.835319],accel_mss,speed_ms,0,blend_radius_m)
  movel([0.265261, -1.342966, -2.575214, -0.794209, 1.570796, 1.836057],accel_mss,speed_ms,0,blend_radius_m)
  movel([0.266136, -1.342591, -2.575461, -0.794337, 1.570796, 1.836932],accel_mss,speed_ms,0,blend_radius_m)
  movel([0.267011, -1.342232, -2.575698, -0.794459, 1.570796, 1.837808],accel_mss,speed_ms,0,blend_radius_m)
  movel([0.267887, -1.341889, -2.575924, -0.794575, 1.570796, 1.838684],accel_mss,speed_ms,0,blend_radius_m)
  movel([0.268764, -1.341565, -2.576138, -0.794686, 1.570796, 1.839560],accel_mss,speed_ms,0,blend_radius_m)
  movel([0.269642, -1.341256, -2.576341, -0.794792, 1.570796, 1.840439],accel_mss,speed_ms,0,blend_radius_m)
  movel([0.270516, -1.340967, -2.576531, -0.794890, 1.570796, 1.841313],accel_mss,speed_ms,0,blend_radius_m)
  movel([0.271393, -1.340694, -2.576711, -0.794984, 1.570796, 1.842189],accel_mss,speed_ms,0,blend_radius_m)
  movel([0.272265, -1.340437, -2.576880, -0.795072, 1.570796, 1.843061],accel_mss,speed_ms,0,blend_radius_m)
  movel([0.273003, -1.340234, -2.577013, -0.795142, 1.570796, 1.843799],accel_mss,speed_ms,0,blend_radius_m)
  movel([0.273733, -1.340049, -2.577135, -0.795205, 1.570796, 1.844529],accel_mss,speed_ms,0,blend_radius_m)
  movel([0.274465, -1.339875, -2.577249, -0.795265, 1.570796, 1.845261],accel_mss,speed_ms,0,blend_radius_m)
  movel([0.275297, -1.339691, -2.577369, -0.795328, 1.570796, 1.846093],accel_mss,speed_ms,0,blend_radius_m)
  movel([0.276127, -1.339518, -2.577483, -0.795388, 1.570796, 1.846923],accel_mss,speed_ms,0,blend_radius_m)
  movel([0.276953, -1.339357, -2.577589, -0.795443, 1.570796, 1.847749],accel_mss,speed_ms,0,blend_radius_m)
  movel([0.278093, -1.339151, -2.577724, -0.795514, 1.570796, 1.848889],accel_mss,speed_ms,0,blend_radius_m)
  movel([0.279230, -1.338962, -2.577848, -0.795579, 1.570796, 1.850026],accel_mss,speed_ms,0,blend_radius_m)
  movel([0.279477, -1.338930, -2.577869, -0.795590, 1.570796, 1.850274],accel_mss,speed_ms,0,blend_radius_m)
  movel([0.279719, -1.338917, -2.577877, -0.795595, 1.570796, 1.850515],accel_mss,speed_ms,0,blend_radius_m)
  movel([0.279954, -1.338919, -2.577876, -0.795594, 1.570796, 1.850750],accel_mss,speed_ms,0,blend_radius_m)
  movel([0.280179, -1.338941, -2.577862, -0.795587, 1.570796, 1.850975],accel_mss,speed_ms,0,blend_radius_m)
  speed_ms = 0.003
  movel([0.280179, -1.342159, -2.579432, -0.790797, 1.570796, 1.850975],accel_mss,speed_ms,0,blend_radius_m)
  speed_ms = 0.007
  movel([0.280440, -1.342192, -2.579411, -0.790786, 1.570796, 1.851236],accel_mss,speed_ms,0,blend_radius_m)
  movel([0.273536, -1.364968, -2.564066, -0.783356, 1.570796, 1.844333],accel_mss,speed_ms,0,blend_radius_m)
  movel([0.270969, -1.373523, -2.558116, -0.780750, 1.570796, 1.841766],accel_mss,speed_ms,0,blend_radius_m)
  movel([0.268811, -1.380723, -2.553029, -0.778636, 1.570796, 1.839607],accel_mss,speed_ms,0,blend_radius_m)
  movel([0.266912, -1.387065, -2.548488, -0.776836, 1.570796, 1.837709],accel_mss,speed_ms,0,blend_radius_m)
  movel([0.266850, -1.387254, -2.548352, -0.776783, 1.570796, 1.837647],accel_mss,speed_ms,0,blend_radius_m)
  movel([0.266777, -1.387443, -2.548216, -0.776730, 1.570796, 1.837573],accel_mss,speed_ms,0,blend_radius_m)
  movel([0.266578, -1.387921, -2.547871, -0.776597, 1.570796, 1.837374],accel_mss,speed_ms,0,blend_radius_m)
  movel([0.264610, -1.388174, -2.547689, -0.776527, 1.570796, 1.835406],accel_mss,speed_ms,0,blend_radius_m)
  movel([0.263843, -1.388265, -2.547623, -0.776501, 1.570796, 1.834640],accel_mss,speed_ms,0,blend_radius_m)
  movel([0.263083, -1.388341, -2.547568, -0.776480, 1.570796, 1.833879],accel_mss,speed_ms,0,blend_radius_m)
  movel([0.262327, -1.388402, -2.547524, -0.776463, 1.570796, 1.833124],accel_mss,speed_ms,0,blend_radius_m)
  movel([0.261578, -1.388447, -2.547491, -0.776451, 1.570796, 1.832375],accel_mss,speed_ms,0,blend_radius_m)
  movel([0.260834, -1.388476, -2.547470, -0.776443, 1.570796, 1.831630],accel_mss,speed_ms,0,blend_radius_m)
  movel([0.260096, -1.388492, -2.547459, -0.776438, 1.570796, 1.830892],accel_mss,speed_ms,0,blend_radius_m)
  movel([0.259365, -1.388490, -2.547460, -0.776439, 1.570796, 1.830161],accel_mss,speed_ms,0,blend_radius_m)
  movel([0.258640, -1.388473, -2.547472, -0.776443, 1.570796, 1.829436],accel_mss,speed_ms,0,blend_radius_m)
  movel([0.257923, -1.388439, -2.547497, -0.776453, 1.570796, 1.828719],accel_mss,speed_ms,0,blend_radius_m)
  movel([0.257213, -1.388392, -2.547531, -0.776466, 1.570796, 1.828010],accel_mss,speed_ms,0,blend_radius_m)
  movel([0.256522, -1.388327, -2.547578, -0.776484, 1.570796, 1.827318],accel_mss,speed_ms,0,blend_radius_m)
  movel([0.255839, -1.388250, -2.547634, -0.776506, 1.570796, 1.826635],accel_mss,speed_ms,0,blend_radius_m)
  movel([0.255166, -1.388154, -2.547702, -0.776532, 1.570796, 1.825962],accel_mss,speed_ms,0,blend_radius_m)
  movel([0.254501, -1.388041, -2.547784, -0.776563, 1.570796, 1.825298],accel_mss,speed_ms,0,blend_radius_m)
  movel([0.253845, -1.387915, -2.547875, -0.776599, 1.570796, 1.824641],accel_mss,speed_ms,0,blend_radius_m)
  movel([0.253200, -1.387773, -2.547978, -0.776638, 1.570796, 1.823996],accel_mss,speed_ms,0,blend_radius_m)
  movel([0.252563, -1.387615, -2.548092, -0.776682, 1.570796, 1.823360],accel_mss,speed_ms,0,blend_radius_m)
  movel([0.251938, -1.387441, -2.548218, -0.776731, 1.570796, 1.822734],accel_mss,speed_ms,0,blend_radius_m)
  movel([0.251323, -1.387251, -2.548354, -0.776784, 1.570796, 1.822119],accel_mss,speed_ms,0,blend_radius_m)
  movel([0.250721, -1.387045, -2.548503, -0.776841, 1.570796, 1.821518],accel_mss,speed_ms,0,blend_radius_m)
  movel([0.250151, -1.386832, -2.548656, -0.776901, 1.570796, 1.820947],accel_mss,speed_ms,0,blend_radius_m)
  movel([0.249594, -1.386603, -2.548821, -0.776965, 1.570796, 1.820390],accel_mss,speed_ms,0,blend_radius_m)
  movel([0.249050, -1.386360, -2.548996, -0.777033, 1.570796, 1.819846],accel_mss,speed_ms,0,blend_radius_m)
  movel([0.248516, -1.386101, -2.549182, -0.777106, 1.570796, 1.819312],accel_mss,speed_ms,0,blend_radius_m)
  movel([0.247995, -1.385828, -2.549379, -0.777182, 1.570796, 1.818792],accel_mss,speed_ms,0,blend_radius_m)
  movel([0.247488, -1.385538, -2.549587, -0.777264, 1.570796, 1.818284],accel_mss,speed_ms,0,blend_radius_m)
  movel([0.246994, -1.385235, -2.549804, -0.777349, 1.570796, 1.817791],accel_mss,speed_ms,0,blend_radius_m)
  movel([0.246515, -1.384916, -2.550033, -0.777439, 1.570796, 1.817311],accel_mss,speed_ms,0,blend_radius_m)
  movel([0.246047, -1.384583, -2.550273, -0.777534, 1.570796, 1.816844],accel_mss,speed_ms,0,blend_radius_m)
  movel([0.245597, -1.384236, -2.550521, -0.777632, 1.570796, 1.816393],accel_mss,speed_ms,0,blend_radius_m)
  movel([0.245219, -1.383924, -2.550745, -0.777721, 1.570796, 1.816016],accel_mss,speed_ms,0,blend_radius_m)
  movel([0.244858, -1.383600, -2.550977, -0.777812, 1.570796, 1.815654],accel_mss,speed_ms,0,blend_radius_m)
  movel([0.244510, -1.383262, -2.551218, -0.777909, 1.570796, 1.815306],accel_mss,speed_ms,0,blend_radius_m)
  movel([0.244175, -1.382913, -2.551468, -0.778008, 1.570796, 1.814972],accel_mss,speed_ms,0,blend_radius_m)
  movel([0.243853, -1.382552, -2.551726, -0.778111, 1.570796, 1.814649],accel_mss,speed_ms,0,blend_radius_m)
  movel([0.243548, -1.382178, -2.551993, -0.778218, 1.570796, 1.814344],accel_mss,speed_ms,0,blend_radius_m)
  movel([0.243259, -1.381790, -2.552270, -0.778329, 1.570796, 1.814056],accel_mss,speed_ms,0,blend_radius_m)
  movel([0.242982, -1.381394, -2.552552, -0.778443, 1.570796, 1.813778],accel_mss,speed_ms,0,blend_radius_m)
  movel([0.242723, -1.380983, -2.552845, -0.778561, 1.570796, 1.813519],accel_mss,speed_ms,0,blend_radius_m)
  movel([0.242476, -1.380563, -2.553143, -0.778683, 1.570796, 1.813273],accel_mss,speed_ms,0,blend_radius_m)
  movel([0.242247, -1.380132, -2.553450, -0.778807, 1.570796, 1.813043],accel_mss,speed_ms,0,blend_radius_m)
  movel([0.242044, -1.379710, -2.553750, -0.778929, 1.570796, 1.812841],accel_mss,speed_ms,0,blend_radius_m)
  movel([0.241857, -1.379274, -2.554059, -0.779056, 1.570796, 1.812653],accel_mss,speed_ms,0,blend_radius_m)
  movel([0.241688, -1.378829, -2.554375, -0.779185, 1.570796, 1.812484],accel_mss,speed_ms,0,blend_radius_m)
  movel([0.241534, -1.378375, -2.554697, -0.779318, 1.570796, 1.812331],accel_mss,speed_ms,0,blend_radius_m)
  movel([0.241400, -1.377909, -2.555026, -0.779454, 1.570796, 1.812197],accel_mss,speed_ms,0,blend_radius_m)
  movel([0.241282, -1.377434, -2.555362, -0.779593, 1.570796, 1.812078],accel_mss,speed_ms,0,blend_radius_m)
  movel([0.241179, -1.376952, -2.555703, -0.779734, 1.570796, 1.811976],accel_mss,speed_ms,0,blend_radius_m)
  movel([0.241096, -1.376458, -2.556051, -0.779879, 1.570796, 1.811892],accel_mss,speed_ms,0,blend_radius_m)
  movel([0.241030, -1.375957, -2.556405, -0.780027, 1.570796, 1.811827],accel_mss,speed_ms,0,blend_radius_m)
  movel([0.240983, -1.375448, -2.556763, -0.780177, 1.570796, 1.811779],accel_mss,speed_ms,0,blend_radius_m)
  movel([0.240954, -1.374939, -2.557122, -0.780328, 1.570796, 1.811750],accel_mss,speed_ms,0,blend_radius_m)
  movel([0.240943, -1.374422, -2.557485, -0.780482, 1.570796, 1.811739],accel_mss,speed_ms,0,blend_radius_m)
  movel([0.240950, -1.373897, -2.557854, -0.780638, 1.570796, 1.811746],accel_mss,speed_ms,0,blend_radius_m)
  movel([0.240977, -1.373365, -2.558227, -0.780797, 1.570796, 1.811774],accel_mss,speed_ms,0,blend_radius_m)
  movel([0.241023, -1.372827, -2.558604, -0.780958, 1.570796, 1.811819],accel_mss,speed_ms,0,blend_radius_m)
  movel([0.241086, -1.372283, -2.558985, -0.781121, 1.570796, 1.811882],accel_mss,speed_ms,0,blend_radius_m)
  movel([0.241165, -1.371737, -2.559367, -0.781285, 1.570796, 1.811962],accel_mss,speed_ms,0,blend_radius_m)
  movel([0.241266, -1.371183, -2.559754, -0.781452, 1.570796, 1.812062],accel_mss,speed_ms,0,blend_radius_m)
  movel([0.241384, -1.370626, -2.560143, -0.781621, 1.570796, 1.812180],accel_mss,speed_ms,0,blend_radius_m)
  movel([0.241521, -1.370065, -2.560534, -0.781791, 1.570796, 1.812317],accel_mss,speed_ms,0,blend_radius_m)
  movel([0.241675, -1.369500, -2.560926, -0.781962, 1.570796, 1.812471],accel_mss,speed_ms,0,blend_radius_m)
  movel([0.241849, -1.368933, -2.561321, -0.782135, 1.570796, 1.812645],accel_mss,speed_ms,0,blend_radius_m)
  movel([0.242040, -1.368364, -2.561716, -0.782309, 1.570796, 1.812836],accel_mss,speed_ms,0,blend_radius_m)
  movel([0.242247, -1.367794, -2.562111, -0.782483, 1.570796, 1.813043],accel_mss,speed_ms,0,blend_radius_m)
  movel([0.242474, -1.367221, -2.562508, -0.782659, 1.570796, 1.813270],accel_mss,speed_ms,0,blend_radius_m)
  movel([0.242718, -1.366647, -2.562906, -0.782836, 1.570796, 1.813514],accel_mss,speed_ms,0,blend_radius_m)
  movel([0.242978, -1.366074, -2.563302, -0.783013, 1.570796, 1.813774],accel_mss,speed_ms,0,blend_radius_m)
  movel([0.243257, -1.365500, -2.563698, -0.783190, 1.570796, 1.814053],accel_mss,speed_ms,0,blend_radius_m)
  movel([0.243552, -1.364927, -2.564094, -0.783368, 1.570796, 1.814348],accel_mss,speed_ms,0,blend_radius_m)
  movel([0.243864, -1.364356, -2.564487, -0.783546, 1.570796, 1.814660],accel_mss,speed_ms,0,blend_radius_m)
  movel([0.244196, -1.363778, -2.564885, -0.783726, 1.570796, 1.814992],accel_mss,speed_ms,0,blend_radius_m)
  movel([0.244544, -1.363205, -2.565279, -0.783905, 1.570796, 1.815340],accel_mss,speed_ms,0,blend_radius_m)
  movel([0.244905, -1.362635, -2.565670, -0.784084, 1.570796, 1.815701],accel_mss,speed_ms,0,blend_radius_m)
  movel([0.245284, -1.362066, -2.566061, -0.784263, 1.570796, 1.816081],accel_mss,speed_ms,0,blend_radius_m)
  movel([0.245678, -1.361499, -2.566449, -0.784441, 1.570796, 1.816475],accel_mss,speed_ms,0,blend_radius_m)
  movel([0.246085, -1.360938, -2.566833, -0.784618, 1.570796, 1.816881],accel_mss,speed_ms,0,blend_radius_m)
  movel([0.246509, -1.360383, -2.567212, -0.784794, 1.570796, 1.817305],accel_mss,speed_ms,0,blend_radius_m)
  movel([0.246944, -1.359830, -2.567590, -0.784969, 1.570796, 1.817741],accel_mss,speed_ms,0,blend_radius_m)
  movel([0.247394, -1.359285, -2.567961, -0.785143, 1.570796, 1.818191],accel_mss,speed_ms,0,blend_radius_m)
  movel([0.247858, -1.358744, -2.568330, -0.785315, 1.570796, 1.818654],accel_mss,speed_ms,0,blend_radius_m)
  movel([0.248368, -1.358172, -2.568719, -0.785498, 1.570796, 1.819164],accel_mss,speed_ms,0,blend_radius_m)
  movel([0.248888, -1.357609, -2.569102, -0.785678, 1.570796, 1.819684],accel_mss,speed_ms,0,blend_radius_m)
  movel([0.249421, -1.357052, -2.569480, -0.785857, 1.570796, 1.820217],accel_mss,speed_ms,0,blend_radius_m)
  movel([0.249964, -1.356502, -2.569853, -0.786034, 1.570796, 1.820760],accel_mss,speed_ms,0,blend_radius_m)
  movel([0.250520, -1.355958, -2.570221, -0.786210, 1.570796, 1.821316],accel_mss,speed_ms,0,blend_radius_m)
  movel([0.251085, -1.355426, -2.570581, -0.786382, 1.570796, 1.821881],accel_mss,speed_ms,0,blend_radius_m)
  movel([0.251663, -1.354899, -2.570938, -0.786553, 1.570796, 1.822460],accel_mss,speed_ms,0,blend_radius_m)
  movel([0.252248, -1.354383, -2.571286, -0.786720, 1.570796, 1.823045],accel_mss,speed_ms,0,blend_radius_m)
  movel([0.252844, -1.353874, -2.571629, -0.786886, 1.570796, 1.823640],accel_mss,speed_ms,0,blend_radius_m)
  movel([0.253467, -1.353363, -2.571973, -0.787052, 1.570796, 1.824263],accel_mss,speed_ms,0,blend_radius_m)
  movel([0.254097, -1.352860, -2.572312, -0.787217, 1.570796, 1.824893],accel_mss,speed_ms,0,blend_radius_m)
  movel([0.254735, -1.352367, -2.572644, -0.787379, 1.570796, 1.825531],accel_mss,speed_ms,0,blend_radius_m)
  movel([0.255380, -1.351883, -2.572969, -0.787537, 1.570796, 1.826176],accel_mss,speed_ms,0,blend_radius_m)
  movel([0.256033, -1.351411, -2.573285, -0.787693, 1.570796, 1.826830],accel_mss,speed_ms,0,blend_radius_m)
  movel([0.256692, -1.350950, -2.573595, -0.787845, 1.570796, 1.827488],accel_mss,speed_ms,0,blend_radius_m)
  movel([0.257360, -1.350498, -2.573897, -0.787994, 1.570796, 1.828157],accel_mss,speed_ms,0,blend_radius_m)
  movel([0.258033, -1.350059, -2.574191, -0.788139, 1.570796, 1.828829],accel_mss,speed_ms,0,blend_radius_m)
  movel([0.258710, -1.349630, -2.574478, -0.788281, 1.570796, 1.829506],accel_mss,speed_ms,0,blend_radius_m)
  movel([0.259422, -1.349196, -2.574768, -0.788425, 1.570796, 1.830218],accel_mss,speed_ms,0,blend_radius_m)
  movel([0.260138, -1.348772, -2.575050, -0.788566, 1.570796, 1.830935],accel_mss,speed_ms,0,blend_radius_m)
  movel([0.260861, -1.348364, -2.575323, -0.788702, 1.570796, 1.831657],accel_mss,speed_ms,0,blend_radius_m)
  movel([0.261586, -1.347966, -2.575588, -0.788835, 1.570796, 1.832382],accel_mss,speed_ms,0,blend_radius_m)
  movel([0.262317, -1.347581, -2.575844, -0.788964, 1.570796, 1.833113],accel_mss,speed_ms,0,blend_radius_m)
  movel([0.263049, -1.347209, -2.576092, -0.789088, 1.570796, 1.833845],accel_mss,speed_ms,0,blend_radius_m)
  movel([0.263783, -1.346851, -2.576330, -0.789208, 1.570796, 1.834579],accel_mss,speed_ms,0,blend_radius_m)
  movel([0.264523, -1.346505, -2.576559, -0.789324, 1.570796, 1.835319],accel_mss,speed_ms,0,blend_radius_m)
  movel([0.265261, -1.346176, -2.576778, -0.789435, 1.570796, 1.836057],accel_mss,speed_ms,0,blend_radius_m)
  movel([0.266136, -1.345802, -2.577026, -0.789561, 1.570796, 1.836932],accel_mss,speed_ms,0,blend_radius_m)
  movel([0.267011, -1.345444, -2.577264, -0.789682, 1.570796, 1.837808],accel_mss,speed_ms,0,blend_radius_m)
  movel([0.267887, -1.345102, -2.577490, -0.789797, 1.570796, 1.838684],accel_mss,speed_ms,0,blend_radius_m)
  movel([0.268764, -1.344778, -2.577704, -0.789907, 1.570796, 1.839560],accel_mss,speed_ms,0,blend_radius_m)
  movel([0.269642, -1.344470, -2.577908, -0.790011, 1.570796, 1.840439],accel_mss,speed_ms,0,blend_radius_m)
  movel([0.270516, -1.344181, -2.578099, -0.790109, 1.570796, 1.841313],accel_mss,speed_ms,0,blend_radius_m)
  movel([0.271393, -1.343909, -2.578279, -0.790201, 1.570796, 1.842189],accel_mss,speed_ms,0,blend_radius_m)
  movel([0.272265, -1.343653, -2.578448, -0.790288, 1.570796, 1.843061],accel_mss,speed_ms,0,blend_radius_m)
  movel([0.273003, -1.343450, -2.578582, -0.790357, 1.570796, 1.843799],accel_mss,speed_ms,0,blend_radius_m)
  movel([0.273733, -1.343265, -2.578704, -0.790420, 1.570796, 1.844529],accel_mss,speed_ms,0,blend_radius_m)
  movel([0.274465, -1.343092, -2.578818, -0.790479, 1.570796, 1.845261],accel_mss,speed_ms,0,blend_radius_m)
  movel([0.275297, -1.342909, -2.578939, -0.790541, 1.570796, 1.846093],accel_mss,speed_ms,0,blend_radius_m)
  movel([0.276127, -1.342736, -2.579053, -0.790600, 1.570796, 1.846923],accel_mss,speed_ms,0,blend_radius_m)
  movel([0.276953, -1.342575, -2.579159, -0.790655, 1.570796, 1.847749],accel_mss,speed_ms,0,blend_radius_m)
  movel([0.278093, -1.342369, -2.579294, -0.790725, 1.570796, 1.848889],accel_mss,speed_ms,0,blend_radius_m)
  movel([0.279230, -1.342181, -2.579418, -0.790790, 1.570796, 1.850026],accel_mss,speed_ms,0,blend_radius_m)
  movel([0.279477, -1.342149, -2.579439, -0.790801, 1.570796, 1.850274],accel_mss,speed_ms,0,blend_radius_m)
  movel([0.279719, -1.342136, -2.579448, -0.790805, 1.570796, 1.850515],accel_mss,speed_ms,0,blend_radius_m)
  movel([0.279954, -1.342138, -2.579447, -0.790804, 1.570796, 1.850750],accel_mss,speed_ms,0,blend_radius_m)
  movel([0.280179, -1.342159, -2.579432, -0.790797, 1.570796, 1.850975],accel_mss,speed_ms,0,blend_radius_m)
  speed_ms = 0.003
  movel([0.280179, -1.329425, -2.573101, -0.809863, 1.570796, 1.850975],accel_mss,speed_ms,0,blend_radius_m)
  speed_ms = 0.01
  movel([0.280179, -1.305078, -2.560060, -0.847250, 1.570796, 1.850975],accel_mss,speed_ms,0,blend_radius_m)
  movel([0.280179, -1.303552, -2.561012, -0.847825, 1.570796, 1.850976],accel_mss,speed_ms,0,blend_radius_m)
  movel([0.280179, -1.327920, -2.574072, -0.810397, 1.570796, 1.850976],accel_mss,speed_ms,0,blend_radius_m)
  speed_ms = 0.003
  movel([0.280179, -1.337445, -2.578840, -0.796104, 1.570796, 1.850976],accel_mss,speed_ms,0,blend_radius_m)
  speed_ms = 0.007
  movel([0.279913, -1.337500, -2.578804, -0.796085, 1.570796, 1.850709],accel_mss,speed_ms,0,blend_radius_m)
  movel([0.279648, -1.337548, -2.578773, -0.796068, 1.570796, 1.850444],accel_mss,speed_ms,0,blend_radius_m)
  movel([0.277856, -1.337840, -2.578582, -0.795967, 1.570796, 1.848653],accel_mss,speed_ms,0,blend_radius_m)
  movel([0.276563, -1.338062, -2.578437, -0.795890, 1.570796, 1.847359],accel_mss,speed_ms,0,blend_radius_m)
  movel([0.275282, -1.338306, -2.578277, -0.795806, 1.570796, 1.846078],accel_mss,speed_ms,0,blend_radius_m)
  movel([0.274151, -1.338544, -2.578121, -0.795724, 1.570796, 1.844947],accel_mss,speed_ms,0,blend_radius_m)
  movel([0.273360, -1.338739, -2.577994, -0.795656, 1.570796, 1.844156],accel_mss,speed_ms,0,blend_radius_m)
  movel([0.271790, -1.339191, -2.577698, -0.795500, 1.570796, 1.842587],accel_mss,speed_ms,0,blend_radius_m)
  movel([0.270212, -1.339694, -2.577368, -0.795327, 1.570796, 1.841008],accel_mss,speed_ms,0,blend_radius_m)
  movel([0.268639, -1.340247, -2.577005, -0.795137, 1.570796, 1.839436],accel_mss,speed_ms,0,blend_radius_m)
  movel([0.267092, -1.340841, -2.576615, -0.794934, 1.570796, 1.837888],accel_mss,speed_ms,0,blend_radius_m)
  movel([0.266404, -1.341114, -2.576435, -0.794840, 1.570796, 1.837200],accel_mss,speed_ms,0,blend_radius_m)
  movel([0.265780, -1.341365, -2.576270, -0.794755, 1.570796, 1.836576],accel_mss,speed_ms,0,blend_radius_m)
  movel([0.265256, -1.341573, -2.576132, -0.794683, 1.570796, 1.836053],accel_mss,speed_ms,0,blend_radius_m)
  movel([0.265076, -1.341645, -2.576085, -0.794659, 1.570796, 1.835873],accel_mss,speed_ms,0,blend_radius_m)
  movel([0.265021, -1.341662, -2.576074, -0.794653, 1.570796, 1.835818],accel_mss,speed_ms,0,blend_radius_m)
  movel([0.265020, -1.341651, -2.576081, -0.794657, 1.570796, 1.835816],accel_mss,speed_ms,0,blend_radius_m)
  movel([0.265096, -1.341602, -2.576114, -0.794674, 1.570796, 1.835892],accel_mss,speed_ms,0,blend_radius_m)
  movel([0.265256, -1.341517, -2.576169, -0.794702, 1.570796, 1.836052],accel_mss,speed_ms,0,blend_radius_m)
  movel([0.265582, -1.341351, -2.576279, -0.794759, 1.570796, 1.836378],accel_mss,speed_ms,0,blend_radius_m)
  movel([0.265910, -1.341194, -2.576382, -0.794813, 1.570796, 1.836706],accel_mss,speed_ms,0,blend_radius_m)
  movel([0.266240, -1.341048, -2.576478, -0.794863, 1.570796, 1.837036],accel_mss,speed_ms,0,blend_radius_m)
  movel([0.266571, -1.340913, -2.576567, -0.794909, 1.570796, 1.837368],accel_mss,speed_ms,0,blend_radius_m)
  movel([0.267667, -1.340489, -2.576846, -0.795054, 1.570796, 1.838463],accel_mss,speed_ms,0,blend_radius_m)
  movel([0.268765, -1.340084, -2.577112, -0.795193, 1.570796, 1.839562],accel_mss,speed_ms,0,blend_radius_m)
  movel([0.269551, -1.339806, -2.577294, -0.795289, 1.570796, 1.840347],accel_mss,speed_ms,0,blend_radius_m)
  movel([0.270337, -1.339535, -2.577472, -0.795382, 1.570796, 1.841133],accel_mss,speed_ms,0,blend_radius_m)
  movel([0.271123, -1.339274, -2.577643, -0.795472, 1.570796, 1.841919],accel_mss,speed_ms,0,blend_radius_m)
  movel([0.271798, -1.339061, -2.577783, -0.795545, 1.570796, 1.842594],accel_mss,speed_ms,0,blend_radius_m)
  movel([0.272471, -1.338859, -2.577915, -0.795615, 1.570796, 1.843268],accel_mss,speed_ms,0,blend_radius_m)
  movel([0.273141, -1.338672, -2.578037, -0.795679, 1.570796, 1.843937],accel_mss,speed_ms,0,blend_radius_m)
  movel([0.273702, -1.338524, -2.578134, -0.795730, 1.570796, 1.844498],accel_mss,speed_ms,0,blend_radius_m)
  movel([0.274262, -1.338387, -2.578224, -0.795778, 1.570796, 1.845058],accel_mss,speed_ms,0,blend_radius_m)
  movel([0.274819, -1.338258, -2.578308, -0.795822, 1.570796, 1.845616],accel_mss,speed_ms,0,blend_radius_m)
  movel([0.275794, -1.338050, -2.578445, -0.795895, 1.570796, 1.846590],accel_mss,speed_ms,0,blend_radius_m)
  movel([0.276766, -1.337858, -2.578570, -0.795961, 1.570796, 1.847563],accel_mss,speed_ms,0,blend_radius_m)
  movel([0.277679, -1.337692, -2.578679, -0.796019, 1.570796, 1.848475],accel_mss,speed_ms,0,blend_radius_m)
  movel([0.278587, -1.337540, -2.578778, -0.796071, 1.570796, 1.849384],accel_mss,speed_ms,0,blend_radius_m)
  movel([0.278988, -1.337484, -2.578814, -0.796090, 1.570796, 1.849784],accel_mss,speed_ms,0,blend_radius_m)
  movel([0.279382, -1.337441, -2.578842, -0.796105, 1.570796, 1.850178],accel_mss,speed_ms,0,blend_radius_m)
  movel([0.279771, -1.337415, -2.578860, -0.796115, 1.570796, 1.850568],accel_mss,speed_ms,0,blend_radius_m)
  movel([0.279984, -1.337406, -2.578866, -0.796118, 1.570796, 1.850780],accel_mss,speed_ms,0,blend_radius_m)
  movel([0.280191, -1.337407, -2.578865, -0.796117, 1.570796, 1.850987],accel_mss,speed_ms,0,blend_radius_m)
  movel([0.280203, -1.337414, -2.578860, -0.796115, 1.570796, 1.850999],accel_mss,speed_ms,0,blend_radius_m)
  movel([0.280197, -1.337433, -2.578848, -0.796108, 1.570796, 1.850993],accel_mss,speed_ms,0,blend_radius_m)
  movel([0.280179, -1.337445, -2.578840, -0.796104, 1.570796, 1.850976],accel_mss,speed_ms,0,blend_radius_m)
  speed_ms = 0.003
  movel([0.280179, -1.340667, -2.580413, -0.791309, 1.570796, 1.850976],accel_mss,speed_ms,0,blend_radius_m)
  speed_ms = 0.007
  movel([0.279913, -1.340722, -2.580377, -0.791290, 1.570796, 1.850709],accel_mss,speed_ms,0,blend_radius_m)
  movel([0.279648, -1.340770, -2.580346, -0.791273, 1.570796, 1.850444],accel_mss,speed_ms,0,blend_radius_m)
  movel([0.277856, -1.341061, -2.580155, -0.791173, 1.570796, 1.848653],accel_mss,speed_ms,0,blend_radius_m)
  movel([0.276563, -1.341282, -2.580009, -0.791097, 1.570796, 1.847359],accel_mss,speed_ms,0,blend_radius_m)
  movel([0.275282, -1.341526, -2.579849, -0.791014, 1.570796, 1.846078],accel_mss,speed_ms,0,blend_radius_m)
  movel([0.274151, -1.341764, -2.579693, -0.790932, 1.570796, 1.844947],accel_mss,speed_ms,0,blend_radius_m)
  movel([0.273360, -1.341958, -2.579565, -0.790866, 1.570796, 1.844156],accel_mss,speed_ms,0,blend_radius_m)
  movel([0.271790, -1.342409, -2.579268, -0.790712, 1.570796, 1.842587],accel_mss,speed_ms,0,blend_radius_m)
  movel([0.270212, -1.342911, -2.578938, -0.790541, 1.570796, 1.841008],accel_mss,speed_ms,0,blend_radius_m)
  movel([0.268639, -1.343463, -2.578573, -0.790353, 1.570796, 1.839436],accel_mss,speed_ms,0,blend_radius_m)
  movel([0.267092, -1.344055, -2.578182, -0.790151, 1.570796, 1.837888],accel_mss,speed_ms,0,blend_radius_m)
  movel([0.266404, -1.344328, -2.578002, -0.790059, 1.570796, 1.837200],accel_mss,speed_ms,0,blend_radius_m)
  movel([0.265780, -1.344578, -2.577837, -0.789974, 1.570796, 1.836576],accel_mss,speed_ms,0,blend_radius_m)
  movel([0.265256, -1.344786, -2.577699, -0.789904, 1.570796, 1.836053],accel_mss,speed_ms,0,blend_radius_m)
  movel([0.265076, -1.344858, -2.577651, -0.789879, 1.570796, 1.835873],accel_mss,speed_ms,0,blend_radius_m)
  movel([0.265021, -1.344875, -2.577640, -0.789874, 1.570796, 1.835818],accel_mss,speed_ms,0,blend_radius_m)
  movel([0.265020, -1.344864, -2.577647, -0.789877, 1.570796, 1.835816],accel_mss,speed_ms,0,blend_radius_m)
  movel([0.265096, -1.344815, -2.577680, -0.789894, 1.570796, 1.835892],accel_mss,speed_ms,0,blend_radius_m)
  movel([0.265256, -1.344730, -2.577736, -0.789923, 1.570796, 1.836052],accel_mss,speed_ms,0,blend_radius_m)
  movel([0.265582, -1.344565, -2.577845, -0.789979, 1.570796, 1.836378],accel_mss,speed_ms,0,blend_radius_m)
  movel([0.265910, -1.344408, -2.577949, -0.790032, 1.570796, 1.836706],accel_mss,speed_ms,0,blend_radius_m)
  movel([0.266240, -1.344262, -2.578045, -0.790081, 1.570796, 1.837036],accel_mss,speed_ms,0,blend_radius_m)
  movel([0.266571, -1.344128, -2.578134, -0.790127, 1.570796, 1.837368],accel_mss,speed_ms,0,blend_radius_m)
  movel([0.267667, -1.343705, -2.578414, -0.790270, 1.570796, 1.838463],accel_mss,speed_ms,0,blend_radius_m)
  movel([0.268765, -1.343300, -2.578681, -0.790408, 1.570796, 1.839562],accel_mss,speed_ms,0,blend_radius_m)
  movel([0.269551, -1.343023, -2.578864, -0.790502, 1.570796, 1.840347],accel_mss,speed_ms,0,blend_radius_m)
  movel([0.270337, -1.342753, -2.579042, -0.790594, 1.570796, 1.841133],accel_mss,speed_ms,0,blend_radius_m)
  movel([0.271123, -1.342492, -2.579214, -0.790683, 1.570796, 1.841919],accel_mss,speed_ms,0,blend_radius_m)
  movel([0.271798, -1.342279, -2.579354, -0.790756, 1.570796, 1.842594],accel_mss,speed_ms,0,blend_radius_m)
  movel([0.272471, -1.342078, -2.579486, -0.790825, 1.570796, 1.843268],accel_mss,speed_ms,0,blend_radius_m)
  movel([0.273141, -1.341892, -2.579608, -0.790889, 1.570796, 1.843937],accel_mss,speed_ms,0,blend_radius_m)
  movel([0.273702, -1.341744, -2.579706, -0.790939, 1.570796, 1.844498],accel_mss,speed_ms,0,blend_radius_m)
  movel([0.274262, -1.341608, -2.579795, -0.790986, 1.570796, 1.845058],accel_mss,speed_ms,0,blend_radius_m)
